(* IEC 61131-3 sources: 2026_Projet_YGO_ExcavatriceDragage/CODE/M_MAIN, 4 files *)

(* ---- GVL_Global.st ---- *)
(* ═══════════════════════════════════════════════════════════════
   🌐 GVL_Global — Variables globales d'utilité générale
   ───────────────────────────────────────────────────────────────
   🎯 Rôle : Horloges et signaux système partagés non persistants.
   📄 Docs : DOC/AF/AF_Partie-02_Architecture_Programme_v3.2.md
   ═══════════════════════════════════════════════════════════════ *)
{attribute 'qualified_only'}
VAR_GLOBAL
    BlinkClock                 : BOOL; // Horloge clignotement système (IHM/diag), rythme réglable GVL_PERSISTENT
END_VAR

(* ---- PRG_04_Treuils_Benne.st ---- *)
(* ═══════════════════════════════════════════════════════════════
   🪝 PRG_04_Treuils_Benne — Commande des Treuils M1 (moteur de retenue) / M2 (moteur Benne), Synchro et Benne
   ───────────────────────────────────────────────────────────────
   ⚙️ Exécuté par la tâche PLC en position 4 (après PRG_03_Modes_Cycle).
   ✅ Arbitre entre les commandes Manuelles (Joystick) et Automatiques (PRG_03_Modes_Cycle).
   📄 Docs : DOC/AF/AF_Partie-10_Fonction_Winch_v2.1.md ; DOC/AF/AF_Partie-10_Fonction_Winch/FB_Bucket_v1.0.md
   ═══════════════════════════════════════════════════════════════ *)

PROGRAM PRG_04_Treuils_Benne

VAR_INPUT
    // === 📥 ENTRÉES PROGRAMME (AUCUNE - PILOTÉ VIA PRG_02 & PRG_03) ===
END_VAR

VAR_OUTPUT
    // === 🚌 BUS INTER-PRG (producteur unique) ===
    Data : ST_WinchInterPrg; // <-- [BUS] Demandes finales, états, sécurités, synchro, benne
END_VAR

VAR
    instWinchSync : FB_WinchSync;
    instBucket   : FB_Bucket;
    // Seuil d'ouverture benne déclarant la fermeture atteinte (FB PUR). Instance PROPRE à
    // PRG_04 : l'arrivée de fermeture est évaluée DANS FB_Bucket, donc sur la mesure du
    // scan même, avant que PRG_04 ne puisse lire ses sorties. Les deux appels portent des
    // entrées identiques au même scan -> même décision, aucun critère dupliqué.
    instCloseThreshold : FB_BucketCloseThreshold;
    ThresholdMeasureValid : BOOL;  // Qualification de la mesure pour la branche seuil (références M1/M2 + défauts + référence benne)
    instSafetyWinchM1 : FB_Safety_Winch;   // Sécurité treuil M1 (SafeStop / permits / PowerCutOff)
    instSafetyWinchM2 : FB_Safety_Winch;
    instWinchM1   : FB_Winch;
    instWinchM2   : FB_Winch;
    // Projection lecture seule des états IHM treuils () : décharge la §8
    // (~250 lignes d'assignations pures) en un FB. Recopie bit-identique des
    // sources → WinchM1State/WinchM2State/WinchM1Safety/WinchM2Safety/CableLimitAscent.
    instWinchStateProjection : FB_WinchStateProjection;
    // Estimateurs bande vitesse réelle : alimentent le garde-fou palier FB_Winch
    // via MeasuredSpeedBand, 1 instance par treuil, mêmes sources que FB_Safety_Winch.
    instWinchLoadEstimatorM1 : FB_WinchLoadEstimator;
    instWinchLoadEstimatorM2 : FB_WinchLoadEstimator;

    // Collecteurs passifs d'apprentissage vitesse par palier : 1 par treuil,
    // écrivent la table RETAIN _WinchSpeedLearnTable {axe x sens x charge/vide x palier}.
    // STRICTEMENT PASSIFS : aucune commande moteur, aucune surveillance survitesse.
    instWinchSpeedLearningM1 : FB_WinchSpeedLearning;
    instWinchSpeedLearningM2 : FB_WinchSpeedLearning;
    // Dérivations des entrées de collecte (charge présente / conditions stables) — voir §6.
    LoadPresentM1 : BOOL;
    LoadPresentM2 : BOOL;
    StableForLearnM1 : BOOL;
    StableForLearnM2 : BOOL;

    // === FB D'ARBITRAGE DE COMMANDE (POO) ===
    instArbM1 : FB_WinchCmdArbitrationM1;  // * [INST] Arbitrage commande treuil M1
    instArbM2 : FB_WinchCmdArbitrationM2;  // * [INST] Arbitrage commande treuil M2
    instArbBucket : FB_BucketCmdArbitration;  // * [INST] Arbitrage commande benne (POO §5)

    // === REQUETES D'AXE ASSEMBLEES AVANT APPEL FB_WINCH ===
    // CODESYS n'accepte pas l'initialiseur de struct anonyme en parametre d'appel :
    // les structs WinchRequest / Sensors / Config sont remplies champ par champ ici.
    ReqM1Winch                   : ST_fbWinch_Req;             // . [LOC] Requête axe M1 (ordre, palier, bornes)
    ReqM2Winch                   : ST_fbWinch_Req;             // . [LOC] Requête axe M2 (ordre, palier, bornes)
    M1WinchSensors               : ST_fbWinch_Sensors;        // . [LOC] Mesures et feedbacks M1
    M2WinchSensors               : ST_fbWinch_Sensors;        // . [LOC] Mesures et feedbacks M2
    M1WinchCfg                   : ST_fbWinch_Cfg;            // . [LOC] Config statique M1 (table paliers, ralentissement)
    M2WinchCfg                   : ST_fbWinch_Cfg;            // . [LOC] Config statique M2 (table paliers, ralentissement)

    // === 📊 STRUCTS INTERNES (publiés via Data) ===
    WinchM1FinalInterlockRequest : ST_WinchFinalInterlockRequest; // . [LOC] Demande finale et interlocks treuil M1
    WinchM2FinalInterlockRequest : ST_WinchFinalInterlockRequest; // . [LOC] Demande finale et interlocks treuil M2
    KoboldContactorCmdArbitrated : BOOL;                         // . [LOC] Ordre contacteur capteur fond Kobold
    WinchM1State                 : ST_WinchState;                // . [LOC] Etat public treuil Retenue M1
    WinchM2State                 : ST_WinchState;                // . [LOC] Etat public treuil Benne M2
    WinchM1Safety                : ST_SafetyWinch;               // . [LOC] Diagnostic et securites treuil M1
    WinchM2Safety                : ST_SafetyWinch;               // . [LOC] Diagnostic et securites treuil M2
    SyncState                    : ST_SyncState;                 // . [LOC] Etat synchronisation treuils M1/M2
    BucketState                  : ST_BucketHMIState;            // . [LOC] Etat de fonctionnement benne
    Benne_IsRoughlyClosed        : BOOL;                         // . [LOC] Benne consideree fermee
    ArmingPermit                 : BOOL;                         // . [LOC] Permission d'armement homme-mort (combiné interlock benne, Option B)

    WinchBothMotionActive : BOOL;
    WinchBothMotionReady         : BOOL;                         // . [LOC] Verrou atomicite demarrage couple : les 2 treuils prets (hors dead-time D18, hors defaut latche)
    WinchBothFinalRequestsCoherent : BOOL;                       // . [LOC] Egalite effective des demandes physiques M1/M2 du scan
    WinchBothFinalStep45Coherent : BOOL;                         // . [LOC] Exception T291-A exacte : descente M1=P4 / M2=P5 en auto AX4..AX7
    WinchBothReqAscent           : BOOL;
    WinchBothReqDescend          : BOOL;
    ManualBottomPositionConfirmed  : BOOL;
    BottomPositionConfirmed        : BOOL;
    CmdBucketCloseArbitrated       : BOOL;

    // Séquencement automatique benne en pilotage both normal --
    // descente uniquement benne ouverte, montée uniquement benne
    // fermée. Distinct de DumpAtTremie/DiveSearch/ExtractionAssist (fonctionnement normal,
    // pas une assistance MAINT_N1/N2 dédiée). Réutilise WinchBothMotionActive/
    // WinchBothMotionDirection (§1 ci-dessus) : déjà exactement "mouvement both
    // demandé" dans les 2 modes (joystick Select=0, ou BtnWinchBothAscent/Descent) — mêmes variables
    // déjà utilisées par instBucket/instDiveSearch/instExtractionAssist.
    WinchBothDiveBucketOpenArmed     : BOOL;  // CmdOpen_IHM déclenché par ce mécanisme (diagnostic IHM)
    WinchBothMotionBlockedByBucket   : BOOL;  // Garde-fou direct -- voir §3
    WinchBothAscentBucketCloseArmed  : BOOL;  // CmdClose_IHM déclenché par ce mécanisme (diagnostic IHM)
    BucketBusyRiseEdge             : R_TRIG; // Détecte le début d'une action benne (Busy monté)
    BucketBusyFallEdge             : F_TRIG; // Détecte la fin d'une action benne (Busy retombé)
    ControlAscentArmedForThisClose : BOOL;   // Mémorise si LA fermeture en cours a été armée par ce mécanisme
    ExtractionControlActive        : BOOL;   // Phase vitesse contrôlée en cours (diagnostic IHM)
    ControlAscentStartM1PosM       : REAL;
    ControlAscentStartM2PosM       : REAL;

    // === ACTION BENNE M2 (bits directionnels, câblés au FB d'arbitrage) ===
    BucketM2ReqAscent  : BOOL;
    BucketM2ReqDescend : BOOL;
    M2AscentPermitApplied : BOOL;
    M2DescendPermitApplied : BOOL;

    // === STRUCTS D'ARBITRAGE (remplis champ par champ, CODESYS refuse l'init anonyme en appel) ===
    ArbIHM     : ST_fbWinchCmdArbitration_IHM;      // . [LOC] Entrées IHM FB d'arbitrage (partagé M1/M2)
    ArbContext : ST_fbWinchCmdArbitration_Context;  // . [LOC] Contexte gating FB d'arbitrage (partagé M1/M2)
    ArbM1Cfg   : ST_fbWinchCmdArbitration_Cfg;      // . [LOC] Config M1 (palier boutons/both)
    ArbM2Cfg   : ST_fbWinchCmdArbitration_Cfg;      // . [LOC] Config M2 (palier boutons/both + override benne)
    ArbBucketIHM     : ST_fbBucketCmdArbitration_IHM;      // . [LOC] Entrées IHM FB d'arbitrage benne
    ArbBucketContext : ST_fbBucketCmdArbitration_Context;  // . [LOC] Contexte gating FB d'arbitrage benne

    M1LogicRunRequest            : BOOL;
    M1LogicReqAscent             : BOOL;
    M1LogicReqDescend            : BOOL;
    M1LogicRequestStepTgt       : INT;   // Palier arbitré M1 (1..5, 0 = arrêt) — consommé par FB_Winch
    M1LogicRequestSpeedCmd_Pct  : REAL;  // Diagnostic % M1 (palier→%, IHM / simu)

    M2LogicRunRequest            : BOOL;
    M2LogicReqAscent             : BOOL;
    M2LogicReqDescend            : BOOL;
    M2LogicRequestStepTgt       : INT;   // Palier arbitré M2 (1..5, 0 = arrêt) — consommé par FB_Winch
    M2LogicRequestSpeedCmd_Pct  : REAL;  // Diagnostic % M2 (palier→%, IHM / simu)

    BottomLimitM1_Active    : REAL;
    BottomLimitM2_Active    : REAL;

    CableLimitAscentM1Reached : BOOL;
    CableLimitAscentM2Reached : BOOL;

    SafeStopM1_Raw          : BOOL;
    SafeStopM2_Raw          : BOOL;
    WinchContactorMismatchLvl1 : BOOL;   // . [LOC] niveau 1 : discordance contacteurs M1/M2 confirmee (amont OU vecteurs finaux) -> SafeStop
    SyncOperationPermit        : BOOL;   // . [LOC] Gate canonique : la surveillance d'ecart M1/M2 (synchro process + MecaE croise) est autorisee. FAUX pendant tout homing / toute manipulation benne.
    BucketActivityHold         : TOF;    // . [LOC] Maintien de la coupure surveillance synchro 4 s APRES la fin d'une action benne (transitoire d'arret treuils : coast + settle codeur -> faux ecart M1/M2)
    SafeStopM1_Active       : BOOL;
    SafeStopM2_Active       : BOOL;
    // Disponibilité de mouvement par axe/sens + conditions de base ArmingPermit
    ArmM1AscentAvail        : BOOL;
    ArmM1DescendAvail       : BOOL;
    ArmM2AscentAvail        : BOOL;
    ArmM2DescendAvail       : BOOL;
    ArmM3TremieAvail        : BOOL;
    ArmM3MaintenanceAvail   : BOOL;
    ArmAnyAxisAvail         : BOOL;
    ArmBucketBusy           : BOOL;
    ArmModeDisabled         : BOOL;
    ArmContactorOff         : BOOL;
    ArmPowerCutOff          : BOOL;
    // Taxonomie permit (D-P1 à D-P11) : SafetyPermit (safety pure), ProcessPermit (process pur),
    // ProcessAndSafetyPermit (= Safety AND Process), EffectivePermit (= couplage synchro).
    SafetyPermitM1_Descend   : BOOL;
    SafetyPermitM2_Descend   : BOOL;
    SafetyPermitM1_Ascent    : BOOL;
    SafetyPermitM2_Ascent    : BOOL;
    ProcessPermitM1_Descend  : BOOL;
    ProcessPermitM2_Descend  : BOOL;
    ProcessPermitM1_Ascent   : BOOL;
    ProcessPermitM2_Ascent   : BOOL;
    ProcessAndSafetyPermitM1_Descend : BOOL;
    ProcessAndSafetyPermitM2_Descend : BOOL;
    ProcessAndSafetyPermitM1_Ascent  : BOOL;
    ProcessAndSafetyPermitM2_Ascent  : BOOL;
    EffectivePermitM1_Descend : BOOL;
    EffectivePermitM2_Descend : BOOL;
    EffectivePermitM1_Ascent  : BOOL;
    EffectivePermitM2_Ascent  : BOOL;
    EffectivePermitBucket_Open  : BOOL;
    EffectivePermitBucket_Close : BOOL;

    // === 🔗 ATOMICITÉ BOTH — états agrégés explicites ===
    // CoupledBoth := couplage atomique M1/M2 indépendant de SyncEnable : actif en
    // synchro classique (anti-télescopage) OU dès qu'un mouvement both est demandé
    // (même si SyncEnable=FALSE en MAINT_N2). Une permission ou un SafeStop d'un
    // treuil bloque alors l'autre : départ jamais isolé.
    CoupledBoth             : BOOL;
    // Diagnostic IHM : Both bloqué + cause priorisée (voir §5).
    BothBlocked             : BOOL;
    BothBlockReason         : E_WinchTraceBlockReason;

    BenneBusyFallEdge     : F_TRIG;

    // Arrêt auto descente sur détection fond Kobold (pilotage normal)
    KoboldAutoStopRiseEdge  : R_TRIG;
    KoboldAutoStopFallEdge  : F_TRIG;
    KoboldImmersionConfirmed: BOOL;
    KoboldBottomTouchLatched: BOOL;
    DescendPermitDiveBucketOpen : BOOL; // mode Dive actif + benne ouverte = descente permise
    // pilotage unitaire M2 "sécurisé" -- bornes ouvert/fermé + palier 1
    ManualBucketLimitsActive : BOOL;
    ManualBucketJogActive    : BOOL; // WinchSel=2 + MAINT : jog benne unitaire M2 (ouv/ferm), indépendant du toggle bornes
    T248BucketJogActive : BOOL; // Phase JOG du séquencement benne-auto couplé (CoupledBucketPhaseLocked) : borne alignée sur l'état franc IsClosed/IsOpen, caduque dès Arbitrated=0
    M2JogApproachOpen        : BOOL; // M2 dans la zone de ralentissement avant l'arrêt ouverture (palier 1)
    M2JogApproachClose       : BOOL; // M2 dans la zone de ralentissement avant l'arrêt fermeture (palier 1)
    SlackCableAscentCapStep1    : BOOL; // mou de câble en récupération -- bride la montée au Palier 1
    BucketNotClosedAscentCapStep1 : BOOL; // benne non fermée à 100% à la montée -- bride la montée au Palier 1

    // Bypass simplifié séquence FB_DiveSearch -- front montant
    // Kobold pendant une descente couplée confirme directement le fond, sans passer par les
    // préconditions strictes de FB_DiveSearch (benne ouverte, DiveStartMin_M, fenêtre immersion).
    // FB_DiveSearch continue de tourner en parallèle (KoboldMeasureEnable toujours câblé
    // dessus) -- ce bypass est un chemin ADDITIONNEL, pas un remplacement.
    BypassKoboldFallEdge       : F_TRIG; // front descendant Kobold
    BypassKoboldBottomTouched  : BOOL;

    SyncMinorDeviation      : BOOL;
    SyncMinorDeviationBlocksUp   : BOOL;
    SyncMinorDeviationBlocksDown : BOOL;
    M2_LimitShift                : REAL;

    EffectiveMaxStepAscent    : INT;
    EffectiveMaxStepDescent  : INT;

    // Plafonds fixes de sécurité en position Maintenance (non réglables IHM).
    MaintenanceMaxStepAscent  : INT;
    MaintenanceMaxStepDescent : INT;

    // Agrégateur de clamp de palier — bornes communes M1=M2 puis M2-propre
    CommonMaxStepAscent   : INT;
    CommonMaxStepDescent : INT;
    CommonMinStepUp   : INT;
    CommonMinStepDown : INT;
    M2MaxStepUp       : INT;
    M2MaxStepDown     : INT;
    M2MinStepUp       : INT;
    M2MinStepDown     : INT;

    // Mémoire scan précédent pour SpeedDelta_Mps (IHM)
    M1_PrevSpeed_Mps : REAL;
    M2_PrevSpeed_Mps : REAL;

    // === MATRICE DE MAINTENANCE N1/N2 (AF-05 §4bis) ===
    // PRG_04 est le producteur unique du bypass EFFECTIF de son axe : FB_Safety_Winch / FB_Winch /
    // FB_Bucket ne connaissent que des booléens déjà gatés, jamais le mode (encapsulation AF03 §2).
    MaintN1 : BOOL;   // . [LOC] Mode MAINT_N1 arbitré (override FDC logiciel momentané)
    MaintN2 : BOOL;   // . [LOC] Mode MAINT_N2 arbitre (secours et pilotage direct contacteurs)
    ExtractionAssistActive : BOOL; // . [LOC] Séquence d'extraction active (mode MAINT + toggle) — gate permis de montée assistée

    // Override du FDC haut LOGICIEL — MAINT_N1, bouton IHM MAINTENU (jamais latché).
    // Le FDC haut CAPTEUR (TopPositionSensor ≈ 8,5 m) n'est JAMAIS ouvert par cet override.
    OverrideTopSoftwareN1M1 : BOOL;
    OverrideTopSoftwareN1M2 : BOOL;

    // Limite haute logicielle active (m) : 7,5 m nominal ➔ 8,5 m (capteur homing haut) sous override.
    TopLimitM1_M : REAL;
    TopLimitM2_M : REAL;

    // Bypass EFFECTIFS de la famille position (= bypass IHM armé, tous modes — dérogation MES 2026).
    // Servent au câblage ET à l'armement du re-homing obligatoire publié vers PRG_03 (PositionLimitOverriddenM1/M2).
    BypassM1TopLimitSwitchEff   : BOOL;
    BypassM1TopLimitSoftwareEff : BOOL;
    BypassM1CableLimitSwitchEff : BOOL;
    BypassM1LimitLegalEff       : BOOL;
    BypassM1MecaDEff            : BOOL;
    BypassM2TopLimitSwitchEff   : BOOL;
    BypassM2TopLimitSoftwareEff : BOOL;
    BypassM2CableLimitSwitchEff : BOOL;
    BypassM2LimitLegalEff       : BOOL;
    BypassM2MecaDEff            : BOOL;

    // Usage effectif d'un override/bypass de position -> arme le re-homing obligatoire (PRG_03).
    PositionLimitOverriddenM1 : BOOL;
    PositionLimitOverriddenM2 : BOOL;
    BrakeForceAllowedM1       : BOOL;
    BrakeForceAllowedM2       : BOOL;
    HomingFreeMoveBlockedN1   : BOOL;

    // 🕵️ Trace de blocage terrain (§8bis) — publiée via Data.TraceM1/M2, consommée FB_TroubleshootingView
    TraceM1               : ST_TraceWinch;        // . [LOC] Trace blocage treuil M1
    TraceM2               : ST_TraceWinch;        // . [LOC] Trace blocage treuil M2
    TraceM1_PrevReason    : E_WinchTraceBlockReason; // . [LOC] Cause précédente M1 (détection de changement)
    TraceM2_PrevReason    : E_WinchTraceBlockReason; // . [LOC] Cause précédente M2 (détection de changement)
END_VAR

{region "🎯 §1 Intention & assistants"}
// === 🪨 §1 INTENTION MAINTENANCE & ASSISTANTS ===

// Consommation de l'intention both continue opérateur (source unique PRG_03, tous modes)
WinchBothMotionActive    := PRG_03_Modes_Cycle.Data.WinchBothIntent.Active;
WinchBothReqAscent  := PRG_03_Modes_Cycle.Data.WinchBothIntent.ReqAscent;
WinchBothReqDescend := PRG_03_Modes_Cycle.Data.WinchBothIntent.ReqDescend;

// Récupération de l'état fond synthétisé par PRG_03
BottomPositionConfirmed := PRG_03_Modes_Cycle.Data.SequenceState.BottomTouchConfirmed;

// MODES DE MAINTENANCE (calculés en tête de scan : consommés dès §2 par instBucket)
// 🚨 DEROGATION MES septembre 2026 (AF-05 §4bis) : les bypass sécurité treuil M1/M2 + benne
// NE SONT PLUS conditionnés au mode. Un bypass IHM armé est effectif dans TOUS les modes
// (y compris SEMI_AUTO / AUTO). Choix opérateur assumé, tracé — voir AF-05 §4bis.
// MAINT_N1 reste utilisé pour l'override momentané du FDC haut logiciel (§5) et l'assistance extraction.
MaintN1 := (PRG_03_Modes_Cycle.Data.Auth.Mode = E_Mode.MAINT_N1);
MaintN2 := (PRG_03_Modes_Cycle.Data.Auth.Mode = E_Mode.MAINT_N2);
// Séquence d'extraction active (mode MAINT + toggle) : gate le permis de montée assistée (§5).
// Le permis lui-même (AscentPermit) est produit par FB_ExtractionAssist et consommé via le contrat benne.
// FB_ExtractionAssist retire (legacy, plus de toggle IHM) : gate desormais toujours ferme.
ExtractionAssistActive := FALSE;

// Jog benne unitaire M2 : joystick dédié M2 (WinchSel=2) en maintenance. Autorise
// l'ouverture (descente M2) hors mode Dive + active la détection passive d'état benne
// dans FB_Bucket. Indépendant du toggle bornes (TglManualBucketLimits).
ManualBucketJogActive := (PRG_03_Modes_Cycle.Data.Auth.JoystickWinchSelectArbitrated = 2)
    AND (PRG_03_Modes_Cycle.Data.Auth.Mode = E_Mode.MAINT_N1 OR PRG_03_Modes_Cycle.Data.Auth.Mode = E_Mode.MAINT_N2);

// Règle absolue en pilotage both normal --
// descente autorisée UNIQUEMENT benne ouverte, montée UNIQUEMENT benne fermée.
// Décision déléguée à FB_BucketCmdArbitration (POO §5) : flags armés + commandes
// arbitrées (ouverture, fermeture, contacteur Kobold). Bit-identique PRG_04 §1/§2.
ArbBucketIHM.BtnOpen  := GVL_IHM.M2TreuilBenne.Bucket.Cmd.BtnOpen;
ArbBucketIHM.BtnClose := GVL_IHM.M2TreuilBenne.Bucket.Cmd.BtnClose;

ArbBucketContext.TglEnableCoupledBucketSequencing := GVL_IHM.Commun.Cfg.TglEnableCoupledBucketSequencing
                                                    AND NOT PRG_02_Acquisition.Data.MachineHoming.Active;
ArbBucketContext.MotionActive   := WinchBothMotionActive;
ArbBucketContext.ReqAscent      := WinchBothReqAscent;
ArbBucketContext.ReqDescend     := WinchBothReqDescend;
ArbBucketContext.BucketIsOpen   := _BucketState.IsOpen;
ArbBucketContext.BucketIsClosed := _BucketState.IsClosed;
ArbBucketContext.CoupledPhaseLocked := PRG_03_Modes_Cycle.Data.Auth.CoupledBucketPhaseLocked;

instArbBucket(
    Enable    := NOT PRG_02_Acquisition.Data.MachineHoming.Active,
    Auth      := PRG_03_Modes_Cycle.Data.Auth,
    ReqBucket := PRG_03_Modes_Cycle.Data.ReqProgram.ReqBucket,
    IHM       := ArbBucketIHM,
    Context   := ArbBucketContext
);
WinchBothDiveBucketOpenArmed    := instArbBucket.WinchBothDiveBucketOpenArmed;
WinchBothAscentBucketCloseArmed := instArbBucket.WinchBothAscentBucketCloseArmed;
CmdBucketCloseArbitrated        := instArbBucket.CmdClose_IHM;
KoboldContactorCmdArbitrated    := instArbBucket.KoboldContactorCmdArbitrated;

{endregion}

{region "🪣 §2 Commande benne"}
// === 🏗️ §2 COMMANDE DU BENNE (FB_Bucket) ===

instBucket(
    Enable              := NOT PRG_03_Modes_Cycle.Data.Auth.InhibitM2,
    Reset               := PRG_07_Supervision.FaultMachineReset_IHM,
    PowerContactorEngaged     := PRG_02_Acquisition.HwIn.Machine.PowerContactorEngaged_DI,
    Mode                := PRG_03_Modes_Cycle.Data.Auth.Mode,
    CmdOpen_IHM         := instArbBucket.CmdOpen_IHM,
    CmdClose_IHM        := CmdBucketCloseArbitrated,
    // 🎛️ Seuil d'ouverture benne déclarant la fermeture atteinte. Réglage lu directement sur
    // GVL_IHM (patron déjà en place dans PRG_04 pour le plafond de montée contrôlée et la
    // distance de contrôle). Aucune copie locale : le FB clôt lui-même la plage, en défense
    // en profondeur.
    CloseReachedOpening_Pct := GVL_IHM.CycleSemiAuto.Cfg.ExtractionStartOpening_Pct,
    HoldAscentP1AfterClose := PRG_03_Modes_Cycle.Data.ReqProgram.ReqBucket.ReqHoldAscentP1AfterClose,
    ReqAscent           := WinchBothReqAscent OR (PRG_03_Modes_Cycle.Data.Auth.Mode = E_Mode.SEMI_AUTO AND PRG_02_Acquisition.Data.Joystick.AxisY.Direction > 0),
    ReqDescend          := WinchBothReqDescend OR (PRG_03_Modes_Cycle.Data.Auth.Mode = E_Mode.SEMI_AUTO AND PRG_02_Acquisition.Data.Joystick.AxisY.Direction < 0),
    EffectivePermitBucket_Open := EffectivePermitBucket_Open,
    EffectivePermitBucket_Close := EffectivePermitBucket_Close,
    CablePosM1          := PRG_02_Acquisition.Data.EncoderM1.Measurement.CablePosM,
    CablePosM2          := PRG_02_Acquisition.Data.EncoderM2.Measurement.CablePosM,
    HomedM1             := PRG_02_Acquisition.Data.EncoderM1.Homed,
    HomedM2             := PRG_02_Acquisition.Data.EncoderM2.Homed,
    HomedAndReliableM1  := PRG_02_Acquisition.Data.EncoderM1.HomedAndReliable,
    HomedAndReliableM2  := PRG_02_Acquisition.Data.EncoderM2.HomedAndReliable,
    HomingSuspectM1     := PRG_02_Acquisition.Data.EncoderM1.HomingSuspect,
    HomingSuspectM2     := PRG_02_Acquisition.Data.EncoderM2.HomingSuspect,
    WinchSelBucket      := (PRG_03_Modes_Cycle.Data.Auth.JoystickWinchSelectArbitrated = 2),
    BucketJogActive     := ManualBucketJogActive,
    ProgramBucketDriveActive := PRG_03_Modes_Cycle.Data.ReqProgram.ReqBucket.ReqOpen
                                OR PRG_03_Modes_Cycle.Data.ReqProgram.ReqBucket.ReqClose
                                OR PRG_03_Modes_Cycle.Data.ReqProgram.ReqBucket.ReqHoldAscentP1AfterClose,
    M1_Busy             := (instWinchM1.StepNumber > 0),
    M2_Busy             := (instWinchM2.StepNumber > 0),
    // Confirmations visuelles N2 : publication et offset benne. Le preset
    // materiel M2 associe est produit independamment dans PRG_02.
    ConfirmOpenPosition  := GVL_IHM.M2TreuilBenne.Bucket.Cmd.BtnConfirmOpenPos,
    ConfirmClosePosition := GVL_IHM.M2TreuilBenne.Bucket.Cmd.BtnConfirmClosePos,
    MachineHomingCommitOpen  := PRG_02_Acquisition.Data.MachineHoming.SetPosBucketOpen,
    MachineHomingCommitClose := PRG_02_Acquisition.Data.MachineHoming.SetPosBucketClose,
    InvalidateRef            := PRG_02_Acquisition.Data.MachineHoming.BucketRefInvalidate,
    MachineHomed := PRG_02_Acquisition.Data.MachineHoming.Homed,
    MachineHomingActive := PRG_02_Acquisition.Data.MachineHoming.Active,
    Config              := _BucketCfgPersist.Config,
    CfgTimeoutDuration     := GVL_IHM.M2TreuilBenne.Bucket.Cfg.CfgTimeoutDuration,
    BucketState        := _BucketState,
    InhibitM1           := PRG_03_Modes_Cycle.Data.Auth.InhibitM1,
    InhibitM2           := PRG_03_Modes_Cycle.Data.Auth.InhibitM2,
    // Bypass benne (n°25 de la matrice) — effectif tous modes si armé (dérogation MES 2026, AF-05 §4bis)
    BypassGlobal        := GVL_IHM.M2TreuilBenne.Bucket.Bypass.Global
);

// Auto-séquencement benne & Dégradation Palier 1
// Si la benne est en cours de fermeture/ouverture (instBucket.Busy), le mouvement couplé attend.
// Si la benne n'est pas fermée (NOT IsClosed) et que instBucket n'est plus occupé (Busy=FALSE),
// toute demande de montée est automatiquement dégradée au Palier 1 (Vitesse lente, voir instWinchM1/M2),
// protégeant ainsi la mécanique même en pilotage unitaire ou si l'auto-séquencement est désactivé.
// 📌 Note d'architecture (lag 1 scan) : M1/M2LogicRequestDirection est consommé ici avant son calcul arbitré
// en §3 (lag d'un cycle automate nominal, toléré et homogène avec les arbitrages Translation/Modes).
WinchBothMotionBlockedByBucket := WinchBothDiveBucketOpenArmed
                                 AND NOT instBucket.Lifecycle.Busy
                                 AND NOT PRG_02_Acquisition.Data.MachineHoming.Active;
BucketNotClosedAscentCapStep1 := NOT ManualBucketJogActive
    AND (M1LogicReqAscent OR M2LogicReqAscent)
    AND NOT instBucket.Lifecycle.Busy
    AND NOT _BucketState.IsClosed;

// === GATE CANONIQUE SURVEILLANCE ECART M1/M2 ===============================================
// REGLE MES : aucun defaut/alarme d'ecart M1/M2 (synchro process, MecaE croise, concordance
// contacteurs) ne doit apparaitre pendant un HOMING (machine ou codeur) ni pendant une
// MANIPULATION BENNE (auto Lifecycle.Busy OU jog unitaire) : dans ces phases M2-M1 varie
// volontairement jusqu'a ~15 m. Ce signal unique coupe la surveillance A LA SOURCE :
//   - instWinchSync.Enable
//   - instSafetyWinchM1/M2.CrossCheckEnable (latch MecaE)
//   - + FB_WinchSync purge ses latch a Enable=FALSE, + FB_Safety_Winch ouvre RefWindow sur
//     NOT CrossCheckEnable (RAZ continue MecaA/E).
// Tempo de RÉACTIVATION : 2 s après la fin d'une action benne (Lifecycle.Busy OU jog
// WinchSel=2), les treuils coastent encore et les codeurs se stabilisent -> l'écart
// serré 0,1 m de FB_WinchSync (SyncDeviationWarn, [SYNC] ErrorID:01) se déclenche à
// tort. Le TOF ne masque QUE FB_WinchSync (gate sur instWinchSync.Enable §4). MecaE
// croisé (tolérance ~2,5 m, absorbe le coast), MecaA et survitesse restent ACTIFS via
// CrossCheckEnable := SyncOperationPermit (inchangé) -> aucun trou de sécurité.
BucketActivityHold(IN := instBucket.Lifecycle.Busy
    OR ManualBucketJogActive
    OR GVL_IHM.M2TreuilBenne.Bucket.Cmd.BtnOpen
    OR GVL_IHM.M2TreuilBenne.Bucket.Cmd.BtnClose
    OR instArbBucket.CmdOpen_IHM
    OR instArbBucket.CmdClose_IHM
    OR PRG_03_Modes_Cycle.Data.ReqProgram.ReqBucket.ReqOpen
    OR PRG_03_Modes_Cycle.Data.ReqProgram.ReqBucket.ReqClose, PT := T#4s);

SyncOperationPermit := PRG_03_Modes_Cycle.Data.Auth.SyncEnable
    AND (PRG_03_Modes_Cycle.Data.Auth.JoystickWinchSelectArbitrated = 0)
    AND NOT PRG_02_Acquisition.Data.MachineHoming.Active
    AND NOT PRG_02_Acquisition.Data.EncoderM1.Measurement.HomingLifecycle.Busy
    AND NOT PRG_02_Acquisition.Data.EncoderM2.Measurement.HomingLifecycle.Busy
    AND NOT instBucket.Lifecycle.Busy
    AND NOT ManualBucketJogActive
    AND NOT GVL_IHM.M2TreuilBenne.Bucket.Cmd.BtnOpen
    AND NOT GVL_IHM.M2TreuilBenne.Bucket.Cmd.BtnClose
    AND NOT instArbBucket.CmdOpen_IHM
    AND NOT instArbBucket.CmdClose_IHM
    AND NOT PRG_03_Modes_Cycle.Data.ReqProgram.ReqBucket.ReqOpen
    AND NOT PRG_03_Modes_Cycle.Data.ReqProgram.ReqBucket.ReqClose
    // Pas de surveillance de synchronisme pendant les phases ou M1/M2 travaillent
    // volontairement de facon dissymetrique : contact fond, retente et fermeture/controle.
    // La surveillance est rearmee a partir de AX12 (montee en charge couplee).
    AND NOT (PRG_03_Modes_Cycle.Data.SequenceState.Step = E_AutoCycleStep.AX8_BOTTOM_CONFIRMED)
    AND NOT (PRG_03_Modes_Cycle.Data.SequenceState.Step = E_AutoCycleStep.AX9_RAISE_OFF_BOTTOM)
    AND NOT (PRG_03_Modes_Cycle.Data.SequenceState.Step = E_AutoCycleStep.AX10_CLOSE_BUCKET)
    AND NOT (PRG_03_Modes_Cycle.Data.SequenceState.Step = E_AutoCycleStep.AX11_CTRL_ASCENT)
    AND instBucket.ActiveOffsetValid;

// En mode récupération (SyncEnable=FALSE), si un mou de câble est détecté (bit3 ErrorId),
// la montée/enroulement est autorisée mais bridée au Palier 1 pour retendre le tambour en sécurité.
// 📌 Note d'architecture (lag 1 scan) : instSafetyWinchM1/M2.ErrorId est consommé ici avant l'exécution du FB
// au §5bis (lag d'un cycle automate nominal, sécurisé en amont par la lecture directe de M2_TensionedCable_DI).
SlackCableAscentCapStep1 := NOT GVL_IHM.Commun.Bypass.SlackCable
    AND NOT PRG_03_Modes_Cycle.Data.Auth.SyncEnable AND (
    ((instSafetyWinchM1.Fault.ErrorId AND 16#0008) <> 16#0000) OR
    ((instSafetyWinchM2.Fault.ErrorId AND 16#0008) <> 16#0000) OR
    (NOT PRG_02_Acquisition.HwIn.Winch.M2_TensionedCable_DI)
);

SyncMinorDeviation := (instWinchSync.Fault.ErrorId AND 16#0001) <> 16#0000;
// 🛡️ Soft-stop synchro : rattrapage directionnel volontaire UNIQUEMENT en
// commande unitaire. En commande BOTH (WinchBothMotionActive), l'écart mineur ne doit
// JAMAIS produire de rattrapage unilatéral d'un seul treuil — il est géré par le clamp
// palier §5ter (les 2 treuils sont bridés à 1) et le seuil critique (SafeStop des 2,
// §5). Donc les drapeaux sync sont coupés dès qu'un mouvement both est demandé.
SyncMinorDeviationBlocksUp   := _SyncSoftStopEnable AND SyncMinorDeviation AND (instWinchSync.SignedDeltaPosM > 0.0) AND NOT WinchBothMotionActive;
SyncMinorDeviationBlocksDown := _SyncSoftStopEnable AND SyncMinorDeviation AND (instWinchSync.SignedDeltaPosM < 0.0) AND NOT WinchBothMotionActive;

IF _CommunCfgPersist.WinchMaxStepAscent <= 0 THEN
    EffectiveMaxStepAscent := 5;
ELSE
    EffectiveMaxStepAscent := _CommunCfgPersist.WinchMaxStepAscent;
END_IF;

IF _CommunCfgPersist.WinchMaxStepDescent <= 0 THEN
    EffectiveMaxStepDescent := 5;
ELSE
    EffectiveMaxStepDescent := _CommunCfgPersist.WinchMaxStepDescent;
END_IF;

{endregion}

{region "🔀 §3 Arbitrage M1/M2"}
// === 🔀 §3 ARBITRAGE CONSIGNES M1 / M2 ===

// ── Arbitrage M1/M2 (FB_WinchCmdArbitrationM1/M2) ──
// Dérivation des bits d'action benne M2 (consommés par les 2 FB d'arbitrage)
BucketM2ReqAscent  := instBucket.M2_ReqAscent;
BucketM2ReqDescend := instBucket.M2_ReqDescend;

// Remplissage des structs d'arbitrage (champ par champ, CODESYS 3.5 refuse l'init anonyme en appel)
ArbIHM.BtnAscentM1           := GVL_IHM.M1TreuilRetenue.Cmd.BtnAscent;
ArbIHM.BtnDescentM1         := GVL_IHM.M1TreuilRetenue.Cmd.BtnDescent;
ArbIHM.BtnAscentM2           := GVL_IHM.M2TreuilBenne.Cmd.BtnAscent;
ArbIHM.BtnDescentM2         := GVL_IHM.M2TreuilBenne.Cmd.BtnDescent;
ArbIHM.BtnWinchBothAscent    := GVL_IHM.Commun.BtnWinchBothAscent;
ArbIHM.BtnWinchBothDescent  := GVL_IHM.Commun.BtnWinchBothDescent;

ArbContext.BucketBusy                     := instBucket.Lifecycle.Busy AND NOT MaintN2;
ArbContext.BucketM2RunRequest             := instBucket.M2_RunRequest AND NOT MaintN2;
ArbContext.BucketM2ReqAscent              := BucketM2ReqAscent;
ArbContext.BucketM2ReqDescend             := BucketM2ReqDescend;
ArbContext.BucketAutoCloseActive          := (PRG_03_Modes_Cycle.Data.Auth.Mode = E_Mode.SEMI_AUTO)
    AND (PRG_03_Modes_Cycle.Data.SequenceState.Step = E_AutoCycleStep.AX10_CLOSE_BUCKET)
    AND PRG_03_Modes_Cycle.Data.ReqProgram.ReqBucket.ReqClose;
ArbContext.BucketHandoffP1Active          := (PRG_03_Modes_Cycle.Data.Auth.Mode = E_Mode.SEMI_AUTO)
    AND (PRG_03_Modes_Cycle.Data.SequenceState.Step = E_AutoCycleStep.AX10B_RACCORDEMENT_P1)
    AND instBucket.CloseReached
    AND PRG_03_Modes_Cycle.Data.ReqProgram.ReqBucket.ReqHoldAscentP1AfterClose;
ArbContext.WinchBothMotionBlockedByBucket := WinchBothMotionBlockedByBucket AND NOT MaintN2;
ArbContext.SyncBlocksAscent                   := SyncMinorDeviationBlocksUp AND NOT MaintN2;
ArbContext.SyncBlocksDescent                 := SyncMinorDeviationBlocksDown AND NOT MaintN2;
// 🔗 Atomicité Both : agrégats consommés par la commande both (§5 calcule
// Both*Permit APRÈS §3 → lag 1 scan assumé au gate d'arbitre, documenté comme les
// autres gates lag-1 de PRG_04 ; l'enforcement même-scan est assuré par le routage
// §6 vers FB_Winch).
ArbContext.M1AscentAllowed  := EffectivePermitM1_Ascent;
ArbContext.M1DescendAllowed := EffectivePermitM1_Descend;
ArbContext.M2AscentAllowed  := EffectivePermitM2_Ascent;
ArbContext.M2DescendAllowed := EffectivePermitM2_Descend;
ArbContext.BothBlock         := BothBlocked;

ArbM1Cfg.BtnStepTgt := 5;
ArbM2Cfg.BtnStepTgt := 5;
ArbM2Cfg.BucketOverrideStepUpTgt   := LIMIT(1, _BucketCfgPersist.Config.MaxStepUp, 5);
ArbM2Cfg.BucketOverrideStepDownTgt := LIMIT(1, _BucketCfgPersist.Config.MaxStepDown, 5);
ArbM2Cfg.BucketAutoMaxStepUp       := LIMIT(1, GVL_IHM.CycleSemiAuto.Cfg.CtrlAscentMaxStep, 2);

// ── Arbitrage M1 (FB_WinchCmdArbitrationM1) ──
instArbM1(
    Enable     := TRUE,
    Joystick   := PRG_02_Acquisition.Data.Joystick,
    Auth       := PRG_03_Modes_Cycle.Data.Auth,
    ReqWinch   := PRG_03_Modes_Cycle.Data.ReqProgram.ReqWinchM1,
    BothIntent := PRG_03_Modes_Cycle.Data.WinchBothIntent,
    IHM        := ArbIHM,
    TglJoystickMaster := GVL_IHM.Modes.Cmd.TglJoystickMaster,
    Context    := ArbContext,
    Cfg        := ArbM1Cfg
);
M1LogicRunRequest := instArbM1.RunRequest;
M1LogicReqAscent  := instArbM1.ReqAscent;
M1LogicReqDescend := instArbM1.ReqDescend;
M1LogicRequestStepTgt := instArbM1.StepTgt;
// Diagnostic % (palier→%) pour IHM / simu — borne haute du palier arbitré.
IF (M1LogicRequestStepTgt >= 1) AND (M1LogicRequestStepTgt <= 5) THEN
    M1LogicRequestSpeedCmd_Pct := _WinchSpeedStepTable.StepThreshold_Pct[M1LogicRequestStepTgt];
ELSE
    M1LogicRequestSpeedCmd_Pct := 0.0;
END_IF;

// ── Arbitrage M2 (FB_WinchCmdArbitrationM2) ──
instArbM2(
    Enable     := TRUE,
    Joystick   := PRG_02_Acquisition.Data.Joystick,
    Auth       := PRG_03_Modes_Cycle.Data.Auth,
    ReqWinch   := PRG_03_Modes_Cycle.Data.ReqProgram.ReqWinchM2,
    BothIntent := PRG_03_Modes_Cycle.Data.WinchBothIntent,
    IHM        := ArbIHM,
    TglJoystickMaster := GVL_IHM.Modes.Cmd.TglJoystickMaster,
    Context    := ArbContext,
    Cfg        := ArbM2Cfg
);
M2LogicRunRequest := instArbM2.RunRequest;
M2LogicReqAscent  := instArbM2.ReqAscent;
M2LogicReqDescend := instArbM2.ReqDescend;
M2LogicRequestStepTgt := instArbM2.StepTgt;

// T248 — HOLD DE TRANSITION : changement de selecteur en cours -> requetes M1/M2 forcees
// a 0 (arret rampe normale) jusqu'a l'arret confirme des 2 treuils. Pas de hand-off en
// mouvement jog<->couple -> supprime l'a-coup. Le mouvement suivant redemarre de zero.
IF PRG_03_Modes_Cycle.Data.Auth.WinchSelTransitionHold THEN
    M1LogicRunRequest := FALSE; M1LogicReqAscent := FALSE; M1LogicReqDescend := FALSE; M1LogicRequestStepTgt := 0;
    M2LogicRunRequest := FALSE; M2LogicReqAscent := FALSE; M2LogicReqDescend := FALSE; M2LogicRequestStepTgt := 0;
END_IF;

// D1/D3/D4/D6 : blocage mouvements libres MAINT_N1 en Step 0 (tant que NOT Homed) + gating directionnel homing
HomingFreeMoveBlockedN1 := MaintN1
                           AND NOT PRG_02_Acquisition.Data.MachineHoming.Homed
                           AND NOT PRG_02_Acquisition.Data.MachineHoming.Active;
IF HomingFreeMoveBlockedN1 THEN
    M1LogicRunRequest := FALSE; M1LogicReqAscent := FALSE; M1LogicReqDescend := FALSE; M1LogicRequestStepTgt := 0;
    M2LogicRunRequest := FALSE; M2LogicReqAscent := FALSE; M2LogicReqDescend := FALSE; M2LogicRequestStepTgt := 0;
ELSIF PRG_02_Acquisition.Data.MachineHoming.Active THEN
    IF PRG_02_Acquisition.Data.MachineHoming.CmdWinchSelect = 2 THEN
        M1LogicRunRequest := FALSE; M1LogicReqAscent := FALSE; M1LogicReqDescend := FALSE; M1LogicRequestStepTgt := 0;
        M2LogicReqAscent  := M2LogicReqAscent  AND PRG_02_Acquisition.Data.MachineHoming.AllowAscent;
        M2LogicReqDescend := M2LogicReqDescend AND PRG_02_Acquisition.Data.MachineHoming.AllowDescend;
        M2LogicRunRequest := M2LogicRunRequest AND (M2LogicReqAscent OR M2LogicReqDescend);
    ELSIF PRG_02_Acquisition.Data.MachineHoming.CmdWinchSelect = 0 THEN
        M1LogicReqAscent  := M1LogicReqAscent  AND PRG_02_Acquisition.Data.MachineHoming.AllowAscent;
        M1LogicReqDescend := M1LogicReqDescend AND PRG_02_Acquisition.Data.MachineHoming.AllowDescend;
        M1LogicRunRequest := M1LogicRunRequest AND (M1LogicReqAscent OR M1LogicReqDescend);
        M2LogicReqAscent  := M2LogicReqAscent  AND PRG_02_Acquisition.Data.MachineHoming.AllowAscent;
        M2LogicReqDescend := M2LogicReqDescend AND PRG_02_Acquisition.Data.MachineHoming.AllowDescend;
        M2LogicRunRequest := M2LogicRunRequest AND (M2LogicReqAscent OR M2LogicReqDescend);
    ELSE
        M1LogicRunRequest := FALSE; M1LogicReqAscent := FALSE; M1LogicReqDescend := FALSE; M1LogicRequestStepTgt := 0;
        M2LogicRunRequest := FALSE; M2LogicReqAscent := FALSE; M2LogicReqDescend := FALSE; M2LogicRequestStepTgt := 0;
    END_IF;
END_IF;
// Diagnostic % (palier→%) pour IHM / simu — borne haute du palier arbitré.
IF (M2LogicRequestStepTgt >= 1) AND (M2LogicRequestStepTgt <= 5) THEN
    M2LogicRequestSpeedCmd_Pct := _WinchSpeedStepTable.StepThreshold_Pct[M2LogicRequestStepTgt];
ELSE
    M2LogicRequestSpeedCmd_Pct := 0.0;
END_IF;

// Front de fin d'action benne (F_TRIG conservé pour §3bis ArmingPermit et extraction control).
// L'arrêt forcé de fin d'action benne est désormais géré en interne par les FB d'arbitrage.
BenneBusyFallEdge(CLK := instBucket.Lifecycle.Busy);

// Après une fermeture benne armée PAR CE mécanisme
// (pas ExtractionAssist, qui a déjà sa propre phase CONTROL_ASCENT), la montée couplée qui
// enchaîne démarre en vitesse contrôlée (palier 1) sur ExtractionControlDistance_M avant de
// repasser en paliers normaux.
BucketBusyRiseEdge(CLK := instBucket.Lifecycle.Busy);
IF BucketBusyRiseEdge.Q THEN
    ControlAscentArmedForThisClose := WinchBothAscentBucketCloseArmed;
END_IF;
IF BucketBusyFallEdge.Q AND ControlAscentArmedForThisClose THEN
    ExtractionControlActive := TRUE;
    ControlAscentStartM1PosM := PRG_02_Acquisition.Data.EncoderM1.Measurement.CablePosM;
    ControlAscentStartM2PosM := PRG_02_Acquisition.Data.EncoderM2.Measurement.CablePosM;
END_IF;
IF ExtractionControlActive THEN
    IF (ABS(PRG_02_Acquisition.Data.EncoderM1.Measurement.CablePosM - ControlAscentStartM1PosM) >= GVL_IHM.CycleSemiAuto.Cfg.ExtractionControlDistance_M)
       AND (ABS(PRG_02_Acquisition.Data.EncoderM2.Measurement.CablePosM - ControlAscentStartM2PosM) >= GVL_IHM.CycleSemiAuto.Cfg.ExtractionControlDistance_M) THEN
        ExtractionControlActive := FALSE;         // Distance de contrôle parcourue : paliers normaux
    ELSIF NOT (WinchBothMotionActive AND WinchBothReqAscent) THEN
        ExtractionControlActive := FALSE;         // Ascending relâchée/interrompue : annule la phase
    END_IF;
END_IF;

{endregion}

{region "🛡️ §3bis ArmingPermit"}
// === 🛡️ §3bis ARMINGPERMIT (général — permis de mouvement) ===
// ArmingPermit = permission d'armement homme-mort (entrée FB_Joystick, consommée PRG_02).
// Règle générale : on ne peut armer QUE si au moins un axe (treuil M1/M2 ou translation M3)
// a un permis de mouvement effectif. Sinon, aucun mouvement n'est possible → armement inutile
// et trompeur (l'opérateur croit pouvoir bouger alors que tout est bloqué).
// Calcul déplacé après §5bis (où EffectivePermitM1/M2_Ascent/Descend sont disponibles).
// Combiné interlock benne conservé : interdit l'armement pendant une action benne
// (instBucket.Lifecycle.Busy) et 1 scan après (BenneBusyFallEdge.Q).
// Polarité positive (NC-100) : TRUE = armement autorisé.
{endregion}

{region "🔄 §4 Synchro M1/M2"}
// === 🔄 §4 SYNCHRONISATION M1 / M2 ===

instWinchSync(
    // Surveillance synchro (ecart position + concordance contacteurs) UNIQUEMENT en
    // pilotage couple. En unitaire M1 ou M2 (JoystickWinchSelectArbitrated <> 0) les
    // deux treuils sont volontairement independants : comparer M1/M2 declencherait un
    // faux ContactorMismatch (M2 commande seul, M1 non) -> SafeStop.
    // Gate canonique SyncOperationPermit (calcule §1) : homing OU benne -> surveillance
    // coupee A LA SOURCE. + ActiveOffsetSettled (transitoire de recalage offset) + inhibitions.
    Enable          := SyncOperationPermit
                        AND instBucket.ActiveOffsetSettled
                        AND NOT BucketActivityHold.Q
                        AND NOT PRG_03_Modes_Cycle.Data.Auth.InhibitM1 AND NOT PRG_03_Modes_Cycle.Data.Auth.InhibitM2,
    Reset           := PRG_07_Supervision.FaultMachineReset_IHM,
    Mode            := PRG_03_Modes_Cycle.Data.Auth.Mode,
    CablePosM1      := PRG_02_Acquisition.Data.EncoderM1.Measurement.CablePosM,
    CablePosM2      := PRG_02_Acquisition.Data.EncoderM2.Measurement.CablePosM,
    HomedAndReliableM1 := PRG_02_Acquisition.Data.EncoderM1.HomedAndReliable,
    HomedAndReliableM2 := PRG_02_Acquisition.Data.EncoderM2.HomedAndReliable,
    SyncEnable      := PRG_03_Modes_Cycle.Data.Auth.SyncEnable,
    CfgSyncToleranceM  := _SyncCfgPersist.CfgSyncTolerance_M,
    CfgSyncCriticalToleranceM := _SyncCfgPersist.CfgSyncCriticalTolerance_M,
    ActiveOffsetM   := instBucket.ActiveOffsetM,
    RelayFwdM1      := instWinchM1.RelayFwd,
    RelayFwdM2      := instWinchM2.RelayFwd,
    RelayRevM1      := instWinchM1.RelayRev,
    RelayRevM2      := instWinchM2.RelayRev,
    Contactor1_M1   := instWinchM1.Contactor1,
    Contactor1_M2   := instWinchM2.Contactor1,
    Contactor2_M1   := instWinchM1.Contactor2,
    Contactor2_M2   := instWinchM2.Contactor2,
    Contactor3_M1   := instWinchM1.Contactor3,
    Contactor3_M2   := instWinchM2.Contactor3,
    Contactor4_M1   := instWinchM1.Contactor4,
    Contactor4_M2   := instWinchM2.Contactor4,
    BypassGlobal    := GVL_IHM.M1M2Sync.Bypass.Global
                       OR GVL_IHM.M1TreuilRetenue.Bypass.Global
                       OR GVL_IHM.M2TreuilBenne.Bypass.Global
                       OR GVL_IHM.M1TreuilRetenue.Bypass.ContactorFeedback
                       OR GVL_IHM.M2TreuilBenne.Bypass.ContactorFeedback
                       OR GVL_IHM.M1TreuilRetenue.Bypass.Safety
                       OR GVL_IHM.M2TreuilBenne.Bypass.Safety
                       OR GVL_IHM.M1TreuilRetenue.Bypass.Process
                       OR GVL_IHM.M2TreuilBenne.Bypass.Process,
    DescentStep45Permit := PRG_03_Modes_Cycle.Data.AutoDiveM1Step4M2Step5Active,
    SpeedStepTable  := _WinchSpeedStepTable
);

// Pas de reconstruction de table M2 : le clamp §5ter (M2MaxStep* := 1) suffit
// — StepNumber ≤ 1 → seuls les états P1 sont commandés.
// M2 consomme directement _WinchSpeedStepTable (table normale).

{endregion}

{region "🔗 §5 Couplage & sécurités"}
// === 🛑 §5 COUPLAGE CROISÉ & SÉCURITÉS ===

// La limite légale (profondeur min. autorisée) doit elle aussi
// bénéficier du ralentissement progressif avant arrêt (comme la limite câble physique), pas juste
// un arrêt sec (DescendPermit). Comme les 2 limites bornent la même
// direction (descente), on alimente FB_Winch.BottomLimitM avec la PLUS RESTRICTIVE des deux
// (MAX de 2 valeurs négatives = celle la moins profonde = atteinte en premier) : le ralentissement
// (FB_Winch §"RALENTISSEMENT AUTOMATIQUE SUR BORDURES") s'enclenche alors sur la bonne limite,
// légale ou câble, sans dupliquer le mécanisme.
// M2 : la limite basse est comparee a CablePosM2 BRUTE cote FB_Winch -> on la decale de
// l'offset benne actif (idem M2_LimitShift cote haut). Benne fermee, M2 a deroule
// ~OffsetCloseM de plus que M1 : sans ce decalage la limite basse M2 se declenche
// ~15 m trop tot (REX MES 2026-09-04). ActiveOffsetM est continu (pente bornee).
IF _CommunCfgPersist.LimitLegalEnabled THEN
    BottomLimitM1_Active := MAX(_WinchM1CfgPersist.CfgCableLimitDescent_M, _CommunCfgPersist.LimitLegalDepthMinAllowed_M);
    BottomLimitM2_Active := MAX(_WinchM2CfgPersist.CfgCableLimitDescent_M, _CommunCfgPersist.LimitLegalDepthMinAllowed_M) + instBucket.ActiveOffsetM;
ELSE
    BottomLimitM1_Active := _WinchM1CfgPersist.CfgCableLimitDescent_M;
    BottomLimitM2_Active := _WinchM2CfgPersist.CfgCableLimitDescent_M + instBucket.ActiveOffsetM;
END_IF;

// 🩺 InputModuleFault (AF06 §3bis) : un module DI TOR hors service rend indisponibles
// les retours frein/thermique/contacteurs/fin de course des DEUX treuils (VH_0800END,
// Local_Digital_IO) — pas de granularité par treuil possible, donc SafeStop des DEUX.
// Perte d'une reference auparavant valide en mouvement : arret controle des
// deux treuils, sans PowerCutOff additionnel. Le cycle libere la demande
// seulement apres le composite d'arret mecanique confirme.
// Discordance contacteurs M1/M2 = niveau 1 (SafeStop) sans masque hexa.
//   - instWinchSync.ContactorMismatch : sur les requetes amont (FB_Winch).
//   - PRG_06_Outputs.Data.ContactorMismatch : sur les vecteurs PHYSIQUES finaux
//     (scan N-1, PRG_06 s'execute apres PRG_04). Escalade -> ExternalSyncEscalation ci-dessous.
WinchContactorMismatchLvl1 := instWinchSync.ContactorMismatch OR PRG_06_Outputs.Data.ContactorMismatch;
SafeStopM1_Raw      := WinchContactorMismatchLvl1 OR instBucket.M1SlipDetected OR PRG_02_Acquisition.Data.InputModules.Fault
                       OR PRG_02_Acquisition.Data.MachineHoming.HomingLoss;
SafeStopM2_Raw      := WinchContactorMismatchLvl1 OR PRG_02_Acquisition.Data.InputModules.Fault
                       OR PRG_02_Acquisition.Data.MachineHoming.HomingLoss;

// Surveillance Kobold descente normale (hors FB_DiveSearch)
// : signal HwIn.Machine.M1_M2_KoboldBottomTouch_DI (même que instDiveSearch §1).
KoboldAutoStopRiseEdge(CLK := PRG_02_Acquisition.HwIn.Machine.M1_M2_KoboldBottomTouch_DI);
KoboldAutoStopFallEdge(CLK := PRG_02_Acquisition.HwIn.Machine.M1_M2_KoboldBottomTouch_DI);

// Levée du verrou au neutre du joystick/boutons ou si toggle désactivé
IF PRG_02_Acquisition.Data.Joystick.AtNeutralXY OR NOT GVL_IHM.Commun.Cfg.TglEnableKoboldAutoStopDescent THEN
    KoboldImmersionConfirmed := FALSE;
    KoboldBottomTouchLatched := FALSE;
END_IF;

// WinchBothMotionActive requis : cette surveillance ne s'arme qu'en pilotage
// BOTH (Select=0), pas en pilotage unitaire M1 (où WinchBothMotionDirection reflète
// quand même l'axe joystick brut).
// Qualification immersion : front montant Kobold dans la fenêtre [ImmersionLower_M..ImmersionUpper_M]
IF GVL_IHM.Commun.Cfg.TglEnableKoboldAutoStopDescent
   AND WinchBothMotionActive
   AND WinchBothReqDescend
   AND _BucketState.IsOpen
   AND KoboldAutoStopRiseEdge.Q THEN
    IF (PRG_02_Acquisition.Data.EncoderM1.Measurement.CablePosM <= GVL_IHM.CycleSemiAuto.Cfg.ImmersionUpper_M)
       AND (PRG_02_Acquisition.Data.EncoderM1.Measurement.CablePosM >= GVL_IHM.CycleSemiAuto.Cfg.ImmersionLower_M)
       AND (PRG_02_Acquisition.Data.EncoderM2.Measurement.CablePosM <= GVL_IHM.CycleSemiAuto.Cfg.ImmersionUpper_M)
       AND (PRG_02_Acquisition.Data.EncoderM2.Measurement.CablePosM >= GVL_IHM.CycleSemiAuto.Cfg.ImmersionLower_M) THEN
        KoboldImmersionConfirmed := TRUE;
    END_IF;
END_IF;

// Détection fond : front descendant Kobold APRÈS immersion confirmée
IF KoboldAutoStopFallEdge.Q AND KoboldImmersionConfirmed THEN
    KoboldBottomTouchLatched := TRUE;
    KoboldImmersionConfirmed := FALSE;
END_IF;

// Autorisation directe et explicite issue de PRG_03 (DiveSearch / Cycle)
DescendPermitDiveBucketOpen := PRG_03_Modes_Cycle.Data.ReqProgram.ReqBucket.DescendPermitDiveBucketOpen;

// Le bypass arrête aussi la descente instantanément, même doctrine que le mécanisme
// KoboldBottomTouchLatched.
// Mode "pilotage unitaire M2 sécurisé" : bornes du JOG MANUEL, portée STRICTE = sélecteur
// arbitré sur M2 seul (Arbitrated=2) + toggle IHM, HORS phase JOG du séquencement benne-auto
// couplé (CoupledBucketPhaseLocked, qui passe aussi par Arbitrated=2 mais possède sa propre
// borne ci-dessous). Ne s'applique
// JAMAIS au pilotage couplé (Arbitrated=0, MAINT ou SEMI_AUTO) : ces mouvements ont leurs
// propres permis process (DescendPermitDiveBucketOpen, séquence auto) et le couplage atomique
// M1/M2 propagerait toute coupure M2 en blocage total des deux treuils. Ne passe PAS par
// instBucket (pas de CloseReq/OpenReq mémorisé, jogging libre) -- bornes directes ouvert/fermé
// (mêmes offsets que FB_Bucket, relatifs à la position réelle de M1) + palier 1 (voir
// instWinchM2 §6 plus bas).
ManualBucketLimitsActive := GVL_IHM.M2TreuilBenne.Bucket.Cmd.TglManualBucketLimits
    AND (PRG_03_Modes_Cycle.Data.Auth.JoystickWinchSelectArbitrated = 2)
    AND NOT PRG_03_Modes_Cycle.Data.Auth.CoupledBucketPhaseLocked
    AND PRG_02_Acquisition.Data.EncoderM1.HomedAndReliable
    AND PRG_02_Acquisition.Data.EncoderM2.HomedAndReliable
    AND NOT (PRG_02_Acquisition.Data.MachineHoming.SoftLimitsOff
             AND PRG_02_Acquisition.Data.MachineHoming.Active);

ProcessPermitM1_Descend := NOT (KoboldBottomTouchLatched OR BypassKoboldBottomTouched) AND DescendPermitDiveBucketOpen;
// Phase JOG du séquencement benne-auto couplé (CoupledBucketPhaseLocked ET Arbitrated=2) :
// borne alignée sur la frontière
// RÉELLE IsClosed/IsOpen (CoherenceLimitM, même seuil que FB_Bucket), jamais sur l'anticipation
// -- sans mouvement pour "coaster" le reste du trajet, une coupure à l'anticipation laisse un
// trou permanent avant l'état franc. Caduque automatiquement dès que Arbitrated repasse à 0
// (phase couplée) : ne bride jamais le mouvement couplé qui suit.
T248BucketJogActive := PRG_03_Modes_Cycle.Data.Auth.CoupledBucketPhaseLocked
    AND (PRG_03_Modes_Cycle.Data.Auth.JoystickWinchSelectArbitrated = 2);
// Ce chemin (pilotage unitaire M2, hors instBucket) applique l'anticipation d'inertie
// OpenAnticipationM/CloseAnticipationM (mêmes que FB_Bucket, réglables IHM) pour couvrir
// aussi le jog unitaire. L'ouverture benne (descente M2) est permise soit par le mode Dive
// (DescendPermitDiveBucketOpen), soit par le jog benne unitaire en maintenance
// (ManualBucketJogActive) — sinon la benne ne pourrait plus s'ouvrir en WinchSel=2.
ProcessPermitM2_Descend := NOT (KoboldBottomTouchLatched OR BypassKoboldBottomTouched)
    AND (DescendPermitDiveBucketOpen OR ManualBucketJogActive)
    AND NOT (ManualBucketLimitsActive AND (PRG_02_Acquisition.Data.EncoderM2.Measurement.CablePosM <= (PRG_02_Acquisition.Data.EncoderM1.Measurement.CablePosM + _BucketCfgPersist.Config.OffsetOpenM + _BucketCfgPersist.Config.OpenAnticipationM)))
    AND NOT (T248BucketJogActive AND (PRG_02_Acquisition.Data.EncoderM2.Measurement.CablePosM <= (PRG_02_Acquisition.Data.EncoderM1.Measurement.CablePosM + _BucketCfgPersist.Config.OffsetOpenM + _BucketCfgPersist.Config.CoherenceLimitM)));

// Permis process de montee : contrat extraction commun aux deux axes.
// M2 conserve l'anticipation de fermeture du pilotage benne unitaire, deja appliquee
// historiquement dans ProcessAndSafetyPermitM2_Ascent (refactor sans changement fonctionnel).
// Meme doctrine que la descente ci-dessus (T248BucketJogActive, CoherenceLimitM).
ProcessPermitM1_Ascent := NOT ExtractionAssistActive
    OR PRG_03_Modes_Cycle.Data.ReqProgram.ReqBucket.AscentPermit;
ProcessPermitM2_Ascent := (NOT ExtractionAssistActive
    OR PRG_03_Modes_Cycle.Data.ReqProgram.ReqBucket.AscentPermit)
    AND NOT (ManualBucketLimitsActive AND (PRG_02_Acquisition.Data.EncoderM2.Measurement.CablePosM >= (PRG_02_Acquisition.Data.EncoderM1.Measurement.CablePosM + _BucketCfgPersist.Config.OffsetCloseM - _BucketCfgPersist.Config.CloseAnticipationM)))
    AND NOT (T248BucketJogActive AND (PRG_02_Acquisition.Data.EncoderM2.Measurement.CablePosM >= (PRG_02_Acquisition.Data.EncoderM1.Measurement.CablePosM + _BucketCfgPersist.Config.OffsetCloseM - _BucketCfgPersist.Config.CoherenceLimitM)));

// Zone de ralentissement jog unitaire M2 : palier 1 forcé dans les JogSlowdownZoneM
// derniers mètres AVANT le point d'arrêt anticipé (Offset ± Anticipation). Le "1 m d'avant"
// est donc calculé sur la cible anticipée, pas sur l'offset brut, et suit tout réglage IHM.
M2JogApproachOpen := ManualBucketJogActive
    AND (PRG_02_Acquisition.Data.EncoderM2.Measurement.CablePosM
         <= (PRG_02_Acquisition.Data.EncoderM1.Measurement.CablePosM
             + _BucketCfgPersist.Config.OffsetOpenM
             + _BucketCfgPersist.Config.OpenAnticipationM
             + _BucketCfgPersist.Config.JogSlowdownZoneM));
M2JogApproachClose := ManualBucketJogActive
    AND (PRG_02_Acquisition.Data.EncoderM2.Measurement.CablePosM
         >= (PRG_02_Acquisition.Data.EncoderM1.Measurement.CablePosM
             + _BucketCfgPersist.Config.OffsetCloseM
             - _BucketCfgPersist.Config.CloseAnticipationM
             - _BucketCfgPersist.Config.JogSlowdownZoneM));

// Decalage de la limite haute logicielle M2 : la benne pend jusqu'a OffsetCloseM sous M1,
// donc en pilotage benne (WinchSel=2) OU si la benne est/va etre fermee, M2 doit avoir la
// marge de montee pour atteindre M1 + OffsetCloseM (pas seulement sa position courante).
// Le latch _BucketState.IsClosed n'est plus stale grace au fix A (§4a efface un latch
// contredit par la mesure). En etat indetermine (jamais latche), le terme WinchSel=2
// garantit quand meme la marge pendant l'operation benne.
// La marge (BIG) est donnee si la benne est/va etre fermee OU des que l'operateur
// SELECTIONNE le mode benne (select joystick BRUT = 2, avant meme l'arbitrage WinchSel) :
// M2 doit pouvoir monter jusqu'a M1 + OffsetCloseM pour fermer. Sinon (benne ouverte,
// M2 suit M1) la limite M2 = celle de M1. Le FDC haut PHYSIQUE reste la barriere dure
// (non bypassable, FB_Safety_Winch:528-531) independamment de cette limite soft.
// Le decalage de la limite M2 = l'offset benne ACTIF, point. Comparer CablePosM2 brute a
// (limite + M2_LimitShift) revient exactement a comparer la position M2 CORRIGEE
// (CablePosM2 - ActiveOffsetM) a la limite nominale - meme reference que M1. L'ancienne
// formule (M1 + OffsetCloseM + 1.5 - CfgCableLimitAscent) suivait M1 avec du retard et
// s'alignait mal selon l'etat benne -> faux declenchement "cable ascent limite" (REX MES
// 2026-09-04 : benne fermee, 15 m deroules, comparaison sur la brute). ActiveOffsetM est
// continu (pente bornee) et suit deja l'ouverture reelle.
M2_LimitShift := instBucket.ActiveOffsetM;

{endregion}

{region "🧮 §5-0 Matrice N1/N2"}
// === 🛡️ §5-0 MATRICE DE MAINTENANCE (AF-05 §4bis) ===
// 🚨 DEROGATION MES septembre 2026 : bypass_effectif := bypass_IHM (armé) — SANS conditionnement
// de mode. Un bypass IHM armé est effectif dans TOUS les modes, SEMI_AUTO et AUTO inclus.
// Écart assumé (Directive Machines / ISO 13849) : traçabilité IHM + doc AF-05 §4bis.
// L'override du FDC haut logiciel reste momentané et propre à MAINT_N1 (§ ci-dessous).

// --- Override FDC haut LOGICIEL (décision Q8) ---------------------------------------------
// MAINT_N1 + bouton IHM MAINTENU ➔ la limite logicielle passe de 7,5 m à la position du capteur
// de homing haut (8,5 m). Relâché ➔ retour à 7,5 m au cycle suivant (aucune mémorisation).
// ⛔ Cet override n'ouvre PAS BypassTopLimitSwitch : le capteur physique haut reste la butée
// dure — si TopPositionSensor retombe, AscentPermit tombe (FB_Safety_Winch §3) ➔ arrêt matériel.
// ⛔ Conditionné à Homed ET NON HomingSuspect : sans référence de position fiable, la butée
// logicielle de FB_Safety_Winch (§3) ET la zone de ralentissement de FB_Winch (§3) sont
// neutralisées — relever la limite dans ce cas ne laisserait QUE le capteur physique comme
// protection, approché à pleine vitesse. Sans référence, il n'y a pas de « dépassement
// contrôlé » : l'override est refusé, seul reste le bypass N2 (acte conscient, tracé).
OverrideTopSoftwareN1M1 := MaintN1
                           AND PRG_02_Acquisition.Data.EncoderM1.Homed
                           AND NOT PRG_02_Acquisition.Data.EncoderM1.HomingSuspect
                           AND GVL_IHM.M1TreuilRetenue.Cmd.BtnOverrideTopSoftware;
OverrideTopSoftwareN1M2 := MaintN1
                           AND PRG_02_Acquisition.Data.EncoderM2.Homed
                           AND NOT PRG_02_Acquisition.Data.EncoderM2.HomingSuspect
                           AND GVL_IHM.M2TreuilBenne.Cmd.BtnOverrideTopSoftware;

// --- Bypass EFFECTIFS de la famille position (individuel OR commun, SANS gate de mode — dérogation MES 2026) ---
BypassM1TopLimitSwitchEff   := (GVL_IHM.M1TreuilRetenue.Bypass.TopLimitSwitch   OR GVL_IHM.Commun.Bypass.TopLimitSwitch);
BypassM1TopLimitSoftwareEff := (GVL_IHM.M1TreuilRetenue.Bypass.TopLimitSoftware OR GVL_IHM.Commun.Bypass.TopLimitSoftware);
BypassM1CableLimitSwitchEff := (GVL_IHM.M1TreuilRetenue.Bypass.CableLimitSwitch OR GVL_IHM.Commun.Bypass.CableLimitSwitch);
BypassM1LimitLegalEff       := (GVL_IHM.M1TreuilRetenue.Bypass.LimitLegal       OR GVL_IHM.Commun.Bypass.LimitLegal);
BypassM1MecaDEff            := GVL_IHM.M1TreuilRetenue.Bypass.MecaD;
BypassM2TopLimitSwitchEff   := (GVL_IHM.M2TreuilBenne.Bypass.TopLimitSwitch      OR GVL_IHM.Commun.Bypass.TopLimitSwitch);
BypassM2TopLimitSoftwareEff := (GVL_IHM.M2TreuilBenne.Bypass.TopLimitSoftware    OR GVL_IHM.Commun.Bypass.TopLimitSoftware);
BypassM2CableLimitSwitchEff := (GVL_IHM.M2TreuilBenne.Bypass.CableLimitSwitch    OR GVL_IHM.Commun.Bypass.CableLimitSwitch);
BypassM2LimitLegalEff       := (GVL_IHM.M2TreuilBenne.Bypass.LimitLegal          OR GVL_IHM.Commun.Bypass.LimitLegal);
BypassM2MecaDEff            := GVL_IHM.M2TreuilBenne.Bypass.MecaD;

// --- Limite haute logicielle active -------------------------------------------------------
// Nominal 7,5 m (CfgCableLimitAscent_M) ; 8,5 m (CfgTopSensorPos_M) sous override N1 momentané
// ou bypass N2 latché du FDC logiciel. M2 conserve son décalage benne (M2_LimitShift) dans les
// deux cas : l'override ne modifie que l'assiette de référence, pas la géométrie M1/M2.
// Le seuil haut nominal est un arrêt immédiat (distance de ralentissement = 0 m).
// En override/bypass MAINT, seul le FDC haut matériel définit la borne : il reste non-bypassable.
TopLimitM1_M := SEL(OverrideTopSoftwareN1M1 OR BypassM1TopLimitSoftwareEff,
                    _CommunCfgPersist.CfgCableLimitAscent_M,
                    _WinchM1CfgPersist.CfgTopSensorPos_M);
TopLimitM2_M := SEL(OverrideTopSoftwareN1M2 OR BypassM2TopLimitSoftwareEff,
                    _CommunCfgPersist.CfgCableLimitAscent_M + M2_LimitShift,
                    _WinchM2CfgPersist.CfgTopSensorPos_M + M2_LimitShift);
// EXEMPTION jog benne seule (WinchSel=2) : la formule ci-dessus, une fois M2_LimitShift
// applique, revient exactement a tester la position REELLE de M1 (M2_raw - ActiveOffsetM
// = M1). Resultat : quand M1 est deja au-dessus de CfgCableLimitAscent_M, fermer/ouvrir
// la benne (M2 seul, M1 IMMOBILE) est bloque par la meme limite que la montee de M1,
// alors que manipuler la benne ne fait jamais monter l'ensemble plus haut que M1 courant
// (REX MES 2026-09-04 : "le treuil ne change pas d'altimetrie en mvt benne"). En jog
// benne pur, on remplace donc la butee ALTITUDE ABSOLUE par une butee GEOMETRIQUE relative
// a M1 courant (OffsetCloseM + marge) : c'est deja le vrai limiteur mecanique de la benne
// (ManualBucketLimitsActive/anticipation, PRG_04 ~710-735). Le FdC haut MATERIEL
// (TopPositionSensor, FB_Safety_Winch) reste une barriere INDEPENDANTE et non affectee.
IF ManualBucketJogActive
   AND PRG_02_Acquisition.Data.EncoderM1.HomedAndReliable
   AND PRG_02_Acquisition.Data.EncoderM2.HomedAndReliable THEN
    TopLimitM2_M := PRG_02_Acquisition.Data.EncoderM1.Measurement.CablePosM
                     + _BucketCfgPersist.Config.OffsetCloseM + 2.0;
ELSIF WinchBothMotionActive AND NOT (OverrideTopSoftwareN1M2 OR BypassM2TopLimitSoftwareEff) THEN
    // En Both (WinchBothMotionActive), M1 est l'autorité nominale de montée et
    // d'arrêt haut. M2 devient un garde-fou dérivé avec marge de tolérance +0.50 m sur le FDC
    // logiciel haut pour éliminer les arrêts prématurés sur benne intermédiaire (réserve TOP >= 1.00 m respectée).
    TopLimitM2_M := _CommunCfgPersist.CfgCableLimitAscent_M + M2_LimitShift + 0.50;
END_IF;

// --- Usage effectif d'un override/bypass de position → re-homing obligatoire ---------------
// Publié vers PRG_03 (rang 03) ➔ FB_Modes arme HomingRequiredMx à la sortie du mode maintenance.
// Famille position : TopLimitSwitch, TopLimitSoftware, CableLimitSwitch, LimitLegal, MecaD
// (+ l'override N1 momentané).
PositionLimitOverriddenM1 := OverrideTopSoftwareN1M1 OR BypassM1TopLimitSwitchEff
                             OR BypassM1TopLimitSoftwareEff OR BypassM1CableLimitSwitchEff
                             OR BypassM1LimitLegalEff OR BypassM1MecaDEff;
PositionLimitOverriddenM2 := OverrideTopSoftwareN1M2 OR BypassM2TopLimitSwitchEff
                             OR BypassM2TopLimitSoftwareEff OR BypassM2CableLimitSwitchEff
                             OR BypassM2LimitLegalEff OR BypassM2MecaDEff;
{endregion}

{region "🛡️ §5bis Sécurité M1/M2"}

// FB_Safety_Winch M1/M2.
// Instancié avant instWinchM1/M2 : MovementCommanded lit RelayFwd/RelayRev du scan précédent
// (même lag 1 scan accepté que M4/Translation, jamais sur Reset/SafeStop/PowerCutOff/sortie finale).
BrakeForceAllowedM1 := MaintN2
    AND PRG_02_Acquisition.HwIn.Machine.EmergencyChainClosed_DI
    AND PRG_02_Acquisition.HwIn.Machine.PowerContactorEngaged_DI
    AND (GVL_IHM.MaintenanceN2.Cmd.BtnBothBrakeRelease OR GVL_IHM.MaintenanceN2.Cmd.BtnM1BrakeRelease);
BrakeForceAllowedM2 := MaintN2
    AND PRG_02_Acquisition.HwIn.Machine.EmergencyChainClosed_DI
    AND PRG_02_Acquisition.HwIn.Machine.PowerContactorEngaged_DI
    AND (GVL_IHM.MaintenanceN2.Cmd.BtnBothBrakeRelease OR GVL_IHM.MaintenanceN2.Cmd.BtnM2BrakeRelease);

instSafetyWinchM1(
    Enable                 := (PRG_03_Modes_Cycle.Data.Auth.Mode <> E_Mode.DISABLE) AND NOT PRG_03_Modes_Cycle.Data.Auth.InhibitM1,
    Reset                  := PRG_07_Supervision.FaultMachineReset_IHM,
    PowerContactorEngaged  := PRG_02_Acquisition.HwIn.Machine.PowerContactorEngaged_DI,
    Mode                   := PRG_03_Modes_Cycle.Data.Auth.Mode,
    SyncEnable             := PRG_03_Modes_Cycle.Data.Auth.SyncEnable,
    CrossCheckEnable       := SyncOperationPermit,
    JoystickOnline         := PRG_02_Acquisition.Data.Network.Joystick.Online,
    JoystickOperational    := PRG_02_Acquisition.Data.Network.Joystick.Operational,
    HeartbeatIhmOk         := GVL_IHM.Commun.HeartbeatIhmOk,
    EncoderAvailable       := PRG_02_Acquisition.Data.EncoderM1.Measurement.EncoderAvailable,
    EncoderFaultBypass     := GVL_IHM.M1TreuilRetenue.Bypass.EncoderFault,
    ThermalFeedback        := NOT PRG_02_Acquisition.HwIn.Winch.M1_ThermalOk_DI,
    BrakeThermalFeedback   := NOT PRG_02_Acquisition.HwIn.Machine.M1_M2_M3_BrakeThermalOk_DI,
    SlackCableDetected     := NOT PRG_02_Acquisition.HwIn.Winch.M2_TensionedCable_DI,
    PhaseRotationOk        := PRG_02_Acquisition.HwIn.Machine.PhaseRotationOk_DI,
    // FB_Safety_Winch attend le contact NC : TRUE = circuit sain / FdC haut libre.
    // FALSE = FdC haut atteint ou rupture de chaîne ; le FB bloque alors la montée.
    TopPositionSensor      := PRG_02_Acquisition.HwIn.Winch.M1M2_TopPositionFree_DI,
    InReferencingMode      := PRG_02_Acquisition.Data.EncoderM1.Measurement.HomingLifecycle.Busy,
    SoftLimitsBypassed     := PRG_02_Acquisition.Data.MachineHoming.SoftLimitsOff
                              AND PRG_02_Acquisition.Data.MachineHoming.Active,
    BrakeForceAllowed      := BrakeForceAllowedM1,
    CablePosM              := PRG_02_Acquisition.Data.EncoderM1.Measurement.CablePosM,
    CfgCableLimitDescentM  := _WinchM1CfgPersist.CfgCableLimitDescent_M,
    LimitLegalReached      := GVL_IHM.Commun.LimitLegalReached,
    ReqAscent              := M1LogicReqAscent,
    ReqDescend             := M1LogicReqDescend,
    MovementCommanded      := instWinchM1.RelayFwd OR instWinchM1.RelayRev,
    Homed                  := PRG_02_Acquisition.Data.EncoderM1.Homed,
    HomingSuspect          := PRG_02_Acquisition.Data.EncoderM1.HomingSuspect,
    TopLimitM              := TopLimitM1_M,
    FwdRevSpeedFeedbackOff := PRG_02_Acquisition.HwIn.Winch.M1_ContactorsReleased_DI,
    BrakeFeedback          := PRG_02_Acquisition.HwIn.Winch.M1_BrakeIsOpen_DI,
    JoystickYNeutral       := (PRG_02_Acquisition.Data.Joystick.AxisY.Direction = 0),
    BenneHoldStillActive   := instBucket.Lifecycle.Busy,
    ExpectedOtherWinchPosM := PRG_02_Acquisition.Data.EncoderM2.Measurement.CablePosM - instBucket.ActiveOffsetM,
    BenneBusy              := instBucket.Lifecycle.Busy,
    OtherWinchInhibited    := PRG_03_Modes_Cycle.Data.Auth.InhibitM2,
    MeasuredSpeedMps       := PRG_02_Acquisition.Data.EncoderM1.Measurement.Speed_Mps,
    MeasuredSpeedSignedMps := PRG_02_Acquisition.Data.EncoderM1.Measurement.SignedSpeed_Mps,
    MeasuredSpeedValid     := PRG_02_Acquisition.Data.EncoderM1.Measurement.SpeedValid,
    SpeedBandMaxMps        := _WinchSpeedConfig.SpeedBandMaxMps[5],
    // Matrice AF-05 §4bis : bypass transmis SANS gate de mode (dérogation MES 2026, tous modes).
    // Le bypass commun reste en OR avec l'individuel (pilotage "both") — câblage d'origine inchangé.
    BypassGlobal           := GVL_IHM.M1TreuilRetenue.Bypass.Global,
    BypassSafety           := GVL_IHM.M1TreuilRetenue.Bypass.Safety,
    BypassProcess          := (GVL_IHM.M1TreuilRetenue.Bypass.Process
                              OR GVL_IHM.Commun.Bypass.SlackCable),
    // OR avec le bypass commun (Commun.Bypass) -- leve la
    // protection sur les 2 treuils simultanement pour le pilotage "both", sans retirer le
    // bypass individuel pour le pilotage a l'unite.
    BypassTopLimitSwitch   := BypassM1TopLimitSwitchEff,
    BypassTopLimitSoftware := BypassM1TopLimitSoftwareEff,
    BypassCableLimitSwitch := BypassM1CableLimitSwitchEff,
    BypassLimitLegal       := BypassM1LimitLegalEff,
    BypassOperatorComm     := GVL_IHM.M1TreuilRetenue.Bypass.OperatorComm,
    BypassPhaseRotation    := GVL_IHM.M1TreuilRetenue.Bypass.PhaseRotation,
    BypassBrakeThermal     := GVL_IHM.M1TreuilRetenue.Bypass.BrakeThermal,
    BypassMotorThermal     := GVL_IHM.M1TreuilRetenue.Bypass.MotorThermal,
    BypassMecaA            := GVL_IHM.M1TreuilRetenue.Bypass.MecaA,
    BypassMecaB            := GVL_IHM.M1TreuilRetenue.Bypass.MecaB,
    BypassMecaC            := GVL_IHM.M1TreuilRetenue.Bypass.MecaC,
    BypassMecaD            := BypassM1MecaDEff,
    BypassMecaE            := GVL_IHM.M1TreuilRetenue.Bypass.MecaE,
    CriticalSyncToleranceM := _WinchCriticalSyncTolerance_M,
    ExternalSyncEscalation := PRG_06_Outputs.Data.ContactorMismatchEscalated,
    TopHardStopLatched     := PRG_06_Outputs.Data.TopHardStopLatched
);

instSafetyWinchM2(
    Enable                 := (PRG_03_Modes_Cycle.Data.Auth.Mode <> E_Mode.DISABLE) AND NOT PRG_03_Modes_Cycle.Data.Auth.InhibitM2,
    Reset                  := PRG_07_Supervision.FaultMachineReset_IHM,
    PowerContactorEngaged  := PRG_02_Acquisition.HwIn.Machine.PowerContactorEngaged_DI,
    Mode                   := PRG_03_Modes_Cycle.Data.Auth.Mode,
    SyncEnable             := PRG_03_Modes_Cycle.Data.Auth.SyncEnable,
    // Ecart critique croise M1/M2 (Meca E, FB_Safety_Winch:354) : gate canonique
    // SyncOperationPermit (homing/benne -> OFF). N'affecte PAS le routage mou-de-cable
    // (:508/:520) qui reste sur SyncEnable brut. Le mouvement couple par boutons-both
    // (WinchBothMotionActive sans WinchSel=0) est un cas residuel -> voir T-tache.
    CrossCheckEnable       := SyncOperationPermit,
    JoystickOnline         := PRG_02_Acquisition.Data.Network.Joystick.Online,
    JoystickOperational    := PRG_02_Acquisition.Data.Network.Joystick.Operational,
    HeartbeatIhmOk         := GVL_IHM.Commun.HeartbeatIhmOk,
    EncoderAvailable       := PRG_02_Acquisition.Data.EncoderM2.Measurement.EncoderAvailable,
    EncoderFaultBypass     := GVL_IHM.M2TreuilBenne.Bypass.EncoderFault,
    ThermalFeedback        := NOT PRG_02_Acquisition.HwIn.Winch.M2_ThermalOk_DI,
    BrakeThermalFeedback   := NOT PRG_02_Acquisition.HwIn.Machine.M1_M2_M3_BrakeThermalOk_DI,
    SlackCableDetected     := NOT PRG_02_Acquisition.HwIn.Winch.M2_TensionedCable_DI,
    PhaseRotationOk        := PRG_02_Acquisition.HwIn.Machine.PhaseRotationOk_DI,
    // Même contact NC que M1 : TRUE = FdC haut libre, FALSE = FdC atteint/chaîne ouverte.
    TopPositionSensor      := PRG_02_Acquisition.HwIn.Winch.M1M2_TopPositionFree_DI,
    InReferencingMode      := PRG_02_Acquisition.Data.EncoderM2.Measurement.HomingLifecycle.Busy,
    SoftLimitsBypassed     := PRG_02_Acquisition.Data.MachineHoming.SoftLimitsOff
                              AND PRG_02_Acquisition.Data.MachineHoming.Active,
    BrakeForceAllowed      := BrakeForceAllowedM2,
    CablePosM              := PRG_02_Acquisition.Data.EncoderM2.Measurement.CablePosM,
    CfgCableLimitDescentM  := _WinchM2CfgPersist.CfgCableLimitDescent_M,
    LimitLegalReached      := GVL_IHM.Commun.LimitLegalReached,
    ReqAscent              := M2LogicReqAscent,
    ReqDescend             := M2LogicReqDescend,
    MovementCommanded      := instWinchM2.RelayFwd OR instWinchM2.RelayRev,
    Homed                  := PRG_02_Acquisition.Data.EncoderM2.Homed,
    HomingSuspect          := PRG_02_Acquisition.Data.EncoderM2.HomingSuspect,
    TopLimitM              := TopLimitM2_M,
    FwdRevSpeedFeedbackOff := PRG_02_Acquisition.HwIn.Winch.M2_ContactorsReleased_DI,
    BrakeFeedback          := PRG_02_Acquisition.HwIn.Winch.M2_BrakeIsOpen_DI,
    JoystickYNeutral       := (PRG_02_Acquisition.Data.Joystick.AxisY.Direction = 0),
    BenneHoldStillActive   := FALSE,
    ExpectedOtherWinchPosM := PRG_02_Acquisition.Data.EncoderM1.Measurement.CablePosM + instBucket.ActiveOffsetM,
    BenneBusy              := instBucket.Lifecycle.Busy,
    OtherWinchInhibited    := PRG_03_Modes_Cycle.Data.Auth.InhibitM1,
    MeasuredSpeedMps       := PRG_02_Acquisition.Data.EncoderM2.Measurement.Speed_Mps,
    MeasuredSpeedSignedMps := PRG_02_Acquisition.Data.EncoderM2.Measurement.SignedSpeed_Mps,
    MeasuredSpeedValid     := PRG_02_Acquisition.Data.EncoderM2.Measurement.SpeedValid,
    SpeedBandMaxMps        := _WinchSpeedConfig.SpeedBandMaxMps[5],
    // Matrice AF-05 §4bis (identique à M1 ci-dessus)
    BypassGlobal           := GVL_IHM.M2TreuilBenne.Bypass.Global,
    BypassSafety           := GVL_IHM.M2TreuilBenne.Bypass.Safety,
    BypassProcess          := (GVL_IHM.M2TreuilBenne.Bypass.Process
                              OR GVL_IHM.Commun.Bypass.SlackCable),
    // OR avec le bypass commun (Commun.Bypass) -- voir M1 ci-dessus
    BypassTopLimitSwitch   := BypassM2TopLimitSwitchEff,
    BypassTopLimitSoftware := BypassM2TopLimitSoftwareEff,
    BypassCableLimitSwitch := BypassM2CableLimitSwitchEff,
    BypassLimitLegal       := BypassM2LimitLegalEff,
    BypassOperatorComm     := GVL_IHM.M2TreuilBenne.Bypass.OperatorComm,
    BypassPhaseRotation    := GVL_IHM.M2TreuilBenne.Bypass.PhaseRotation,
    BypassBrakeThermal     := GVL_IHM.M2TreuilBenne.Bypass.BrakeThermal,
    BypassMotorThermal     := GVL_IHM.M2TreuilBenne.Bypass.MotorThermal,
    BypassMecaA            := GVL_IHM.M2TreuilBenne.Bypass.MecaA,
    BypassMecaB            := GVL_IHM.M2TreuilBenne.Bypass.MecaB,
    BypassMecaC            := GVL_IHM.M2TreuilBenne.Bypass.MecaC,
    BypassMecaD            := BypassM2MecaDEff,
    BypassMecaE            := GVL_IHM.M2TreuilBenne.Bypass.MecaE,
    CriticalSyncToleranceM := _WinchCriticalSyncTolerance_M,
    ExternalSyncEscalation := PRG_06_Outputs.Data.ContactorMismatchEscalated,
    TopHardStopLatched     := PRG_06_Outputs.Data.TopHardStopLatched
);

SafeStopM1_Raw := SafeStopM1_Raw OR instSafetyWinchM1.SafeStop;
SafeStopM2_Raw := SafeStopM2_Raw OR instSafetyWinchM2.SafeStop;
// SafetyPermit = sorties FB_Safety_Winch (safety pure)
SafetyPermitM1_Descend := instSafetyWinchM1.DescendPermit;
SafetyPermitM2_Descend := instSafetyWinchM2.DescendPermit;
SafetyPermitM1_Ascent  := instSafetyWinchM1.AscentPermit;
SafetyPermitM2_Ascent  := instSafetyWinchM2.AscentPermit;
// ProcessAndSafetyPermit = Safety AND Process (ex _Raw)
ProcessAndSafetyPermitM1_Descend := ProcessPermitM1_Descend AND SafetyPermitM1_Descend;
ProcessAndSafetyPermitM2_Descend := ProcessPermitM2_Descend AND SafetyPermitM2_Descend;

// Mode "vidage à la trémie" : descente M1 interdite tant que M3 n'est pas à P1 (travail)
// ou en position Maintenance -- verrouille la descente-treuil (payout cable reel) / la
// translation, pour se rapprocher d'un enchaînement automatique sûr.
// M2 EXEMPTE quand seule la benne bouge (jog unitaire WinchSel=2 ou programme benne) :
// ouvrir/fermer la benne (M2 seul, M1 immobile) N'EST PAS une descente treuil verticale
// -> ça doit rester possible a la Tremie (design d'origine : "a la Tremie, seul open/close
// benne permis"). Sans cette exemption, EffectivePermitBucket_Open/Close (cable sur
// EffectivePermitM2_Descend/Ascent, ligne ~1004) heritait du meme verrou par accident de
// cablage -> ouverture benne bloquee a la Tremie (REX MES 2026-09-04).
// Décision et calcul centralisés dans PRG_03_Modes_Cycle.Data.SequenceState.WinchDescentAuth_M3
IF NOT PRG_03_Modes_Cycle.Data.SequenceState.WinchDescentAuth_M3 THEN
    ProcessAndSafetyPermitM1_Descend := FALSE;
    IF NOT (ManualBucketJogActive
            OR PRG_03_Modes_Cycle.Data.ReqProgram.ReqBucket.ReqOpen
            OR PRG_03_Modes_Cycle.Data.ReqProgram.ReqBucket.ReqClose) THEN
        ProcessAndSafetyPermitM2_Descend := FALSE;
    END_IF;
END_IF;
// Permis de montée assistée : consommé depuis FB_ExtractionAssist (via le contrat benne).
// Hors extraction (NOT ExtractionAssistActive), la montée reste libre ; pendant l'extraction,
// la montée n'est autorisée que si l'assistant la délivre (AscentPermit, qui intègre les
// conditions process AscentControlSafe/AscentNominalSafe). Polarité fail-safe (TRUE = autorisé).
ProcessAndSafetyPermitM1_Ascent := ProcessPermitM1_Ascent AND SafetyPermitM1_Ascent;
ProcessAndSafetyPermitM2_Ascent := ProcessPermitM2_Ascent AND SafetyPermitM2_Ascent;

// 🔗 Couplage atomique M1/M2 : indépendant de SyncEnable. Actif en synchro
// classique (anti-télescopage) OU dès qu'un mouvement both est demandé — même si
// SyncEnable=FALSE (ex. MAINT_N2). Permet qu'une permission ou un SafeStop d'un
// treuil bloque l'autre : départ jamais isolé. WinchBothMotionActive est défini en
// §1 (disponible avant §5).
CoupledBoth := instWinchSync.SyncActive OR WinchBothMotionActive;

SafeStopM1_Active := SafeStopM1_Raw OR (CoupledBoth AND SafeStopM2_Raw);
SafeStopM2_Active := SafeStopM2_Raw OR (CoupledBoth AND SafeStopM1_Raw);
// EffectivePermit = ProcessAndSafetyPermit combine au couplage synchro (anti-télescopage)
// ET gaté par NOT SafeStop (défauts thermique/phase/codeur/méca) : le permit reflète « prêt à
// fonctionner », aligné sur M3 (PRG_05 §1ter). SafeStopM1/M2_Active agrège déjà le couplage
// synchro (SafeStop de l'autre treuil pendant SyncActive) — cohérent avec l'anti-télescopage.
EffectivePermitM1_Descend := ProcessAndSafetyPermitM1_Descend AND NOT SafeStopM1_Active AND (NOT CoupledBoth OR ProcessAndSafetyPermitM2_Descend);
EffectivePermitM2_Descend := ProcessAndSafetyPermitM2_Descend AND NOT SafeStopM2_Active AND (NOT CoupledBoth OR ProcessAndSafetyPermitM1_Descend);
EffectivePermitM1_Ascent  := ProcessAndSafetyPermitM1_Ascent  AND NOT SafeStopM1_Active AND (NOT CoupledBoth OR ProcessAndSafetyPermitM2_Ascent);
EffectivePermitM2_Ascent  := ProcessAndSafetyPermitM2_Ascent  AND NOT SafeStopM2_Active AND (NOT CoupledBoth OR ProcessAndSafetyPermitM1_Ascent);

// Mode secours MAINT_N2 : pilotage direct inconditionnel des contacteurs M1/M2 (ensemble ou separement)
// sous la seule reserve de la chaine AU physique fermee (PowerContactorEngaged_DI) et du capteur
// mecanique haut (TopPositionFree_DI, sauf bypass explicite).
IF MaintN2 THEN
    SafeStopM1_Active := NOT PRG_02_Acquisition.HwIn.Machine.PowerContactorEngaged_DI;
    SafeStopM2_Active := NOT PRG_02_Acquisition.HwIn.Machine.PowerContactorEngaged_DI;
    EffectivePermitM1_Descend := PRG_02_Acquisition.HwIn.Machine.PowerContactorEngaged_DI;
    EffectivePermitM2_Descend := PRG_02_Acquisition.HwIn.Machine.PowerContactorEngaged_DI;
    EffectivePermitM1_Ascent  := PRG_02_Acquisition.HwIn.Machine.PowerContactorEngaged_DI
                                 AND ((PRG_02_Acquisition.HwIn.Winch.M1M2_TopPositionFree_DI
                                       AND NOT PRG_06_Outputs.Data.TopHardStopLatched)
                                      OR BypassM1TopLimitSwitchEff
                                      OR GVL_IHM.M1TreuilRetenue.Bypass.Global);
    EffectivePermitM2_Ascent  := PRG_02_Acquisition.HwIn.Machine.PowerContactorEngaged_DI
                                 AND ((PRG_02_Acquisition.HwIn.Winch.M1M2_TopPositionFree_DI
                                       AND NOT PRG_06_Outputs.Data.TopHardStopLatched)
                                      OR BypassM2TopLimitSwitchEff
                                      OR GVL_IHM.M2TreuilBenne.Bypass.Global);
END_IF;

// Si un cycle homing machine est actif (en N1 ou N2), appliquer ses permis par etape
IF HomingFreeMoveBlockedN1 THEN
    EffectivePermitM1_Ascent  := FALSE;
    EffectivePermitM1_Descend := FALSE;
    EffectivePermitM2_Ascent  := FALSE;
    EffectivePermitM2_Descend := FALSE;
ELSIF PRG_02_Acquisition.Data.MachineHoming.Active THEN
    IF PRG_02_Acquisition.Data.MachineHoming.CmdWinchSelect = 2 THEN
        EffectivePermitM1_Ascent  := FALSE;
        EffectivePermitM1_Descend := FALSE;
        EffectivePermitM2_Ascent  := EffectivePermitM2_Ascent  AND PRG_02_Acquisition.Data.MachineHoming.AllowAscent;
        EffectivePermitM2_Descend := EffectivePermitM2_Descend AND PRG_02_Acquisition.Data.MachineHoming.AllowDescend;
    ELSIF PRG_02_Acquisition.Data.MachineHoming.CmdWinchSelect = 0 THEN
        EffectivePermitM1_Ascent  := EffectivePermitM1_Ascent  AND PRG_02_Acquisition.Data.MachineHoming.AllowAscent;
        EffectivePermitM1_Descend := EffectivePermitM1_Descend AND PRG_02_Acquisition.Data.MachineHoming.AllowDescend;
        EffectivePermitM2_Ascent  := EffectivePermitM2_Ascent  AND PRG_02_Acquisition.Data.MachineHoming.AllowAscent;
        EffectivePermitM2_Descend := EffectivePermitM2_Descend AND PRG_02_Acquisition.Data.MachineHoming.AllowDescend;
    ELSE
        EffectivePermitM1_Ascent  := FALSE;
        EffectivePermitM1_Descend := FALSE;
        EffectivePermitM2_Ascent  := FALSE;
        EffectivePermitM2_Descend := FALSE;
    END_IF;
END_IF;

// Permis canoniques benne : ouverture = M2 vers le bas, fermeture = M2 vers le haut.
// Les fins de course benne restent des faits fonctionnels distincts des limites treuil.
EffectivePermitBucket_Open := EffectivePermitM2_Descend
    AND PRG_02_Acquisition.Data.EncoderM1.Homed
    AND PRG_02_Acquisition.Data.EncoderM2.Homed
    AND (instBucket.Lifecycle.Busy OR NOT _BucketState.IsOpen)
    AND NOT instBucket.Fault.Error;
EffectivePermitBucket_Close := EffectivePermitM2_Ascent
    AND PRG_02_Acquisition.Data.EncoderM1.Homed
    AND PRG_02_Acquisition.Data.EncoderM2.Homed
    AND (instBucket.Lifecycle.Busy OR NOT _BucketState.IsClosed)
    AND NOT instBucket.Fault.Error;

// Défense en profondeur benne : le permis directionnel benne est appliqué au
// même scan aux deux niveaux M2, uniquement lorsque FB_Bucket est producteur.
M2AscentPermitApplied := EffectivePermitM2_Ascent
    AND (NOT instBucket.M2_RunRequest OR EffectivePermitBucket_Close);
M2DescendPermitApplied := EffectivePermitM2_Descend
    AND (NOT instBucket.M2_RunRequest OR EffectivePermitBucket_Open);

// 🔗 Agrégats Both : permis communs consommés par la commande both.
// = AND des 4 permits effectifs. Chaque axe garde sa vérité propre
// (EffectivePermitM*_*) ; en commande both, seul l'agrégat est consommé (§6),
// garantissant "les 2 treuils partent ensemble, ou aucun".

// 📉 Diagnostic IHM — cause priorisée du blocage Both (lecture seule, NC-100).
// N'a AUCUN effet de conduite : l'arrêt est porté par Both*Permit (§6, consommé par les
// 2 FB_Winch) et la défense en profondeur par la barrière finale (FB_WinchOutputInterlock,
// coupe par PermitFinalBlocked). Ordre : cause la plus grave gagne.
IF NOT WinchBothMotionActive THEN
    BothBlocked             := FALSE;
    BothBlockReason         := E_WinchTraceBlockReason.NONE;
ELSIF NOT ((WinchBothReqAscent AND EffectivePermitM1_Ascent AND EffectivePermitM2_Ascent)
        OR (WinchBothReqDescend AND EffectivePermitM1_Descend AND EffectivePermitM2_Descend)) THEN
    BothBlocked             := TRUE;
    BothBlockReason         := E_WinchTraceBlockReason.COUPLING_BLOCKED;
ELSE
    BothBlocked             := FALSE;
    BothBlockReason         := E_WinchTraceBlockReason.NONE;
END_IF;

// 🛡️ ArmingPermit : armer HONNETEMENT, seulement si au moins une action
// selectionnee peut REELLEMENT partir. Disponibilite par axe x sens + motif de
// blocage decode pour l'IHM / troubleshooting. Reprise apres perte = nouveau front
// homme-mort global (FB_Joystick : IF NOT ArmingPermit -> desarme le geste entier).
// EffectivePermitM*_* couvre deja process + safety + NOT SafeStop de cet axe +
// verif couplage ; on ajoute NOT Fault.Latched (faute finale) et, pour M3, le
// permis effectif directionnel + SafeStop/PowerCutOff M3 (bus PRG_05, lag 1 scan).
ArmM1AscentAvail  := EffectivePermitM1_Ascent  AND (MaintN2 OR NOT instSafetyWinchM1.Fault.Latched);
ArmM1DescendAvail := EffectivePermitM1_Descend AND (MaintN2 OR NOT instSafetyWinchM1.Fault.Latched);
ArmM2AscentAvail  := EffectivePermitM2_Ascent  AND (MaintN2 OR NOT instSafetyWinchM2.Fault.Latched);
ArmM2DescendAvail := EffectivePermitM2_Descend AND (MaintN2 OR NOT instSafetyWinchM2.Fault.Latched);
ArmM3TremieAvail  := PRG_05_Translation.Data.TranslationFinalInterlockRequest.EffectivePermitM3_Tremie
                     AND NOT PRG_05_Translation.Data.TranslationSafety.SafeStop
                     AND NOT PRG_05_Translation.Data.TranslationSafety.PowerCutOff;
ArmM3MaintenanceAvail := PRG_05_Translation.Data.TranslationFinalInterlockRequest.EffectivePermitM3_Maintenance
                     AND NOT PRG_05_Translation.Data.TranslationSafety.SafeStop
                     AND NOT PRG_05_Translation.Data.TranslationSafety.PowerCutOff;

ArmAnyAxisAvail := ArmM1AscentAvail OR ArmM1DescendAvail
               OR ArmM2AscentAvail OR ArmM2DescendAvail
               OR ArmM3TremieAvail OR ArmM3MaintenanceAvail;

// Conditions de base (AC1) — priorite decroissante pour le motif.
// En SEMI_AUTO ou lors d'une commande benne programme (AX3_OPEN_BUCKET / vidage), l'operateur
// doit pouvoir armer l'homme-mort (DeadmanArmed) pour autoriser le mouvement benne !
ArmBucketBusy := (instBucket.Lifecycle.Busy OR BenneBusyFallEdge.Q)
                 AND NOT MaintN2
                 AND NOT PRG_02_Acquisition.Data.MachineHoming.Active
                 AND (PRG_03_Modes_Cycle.Data.Auth.Mode <> E_Mode.SEMI_AUTO)
                 AND NOT PRG_03_Modes_Cycle.Data.ReqProgram.ReqBucket.ReqOpen
                 AND NOT PRG_03_Modes_Cycle.Data.ReqProgram.ReqBucket.ReqClose;
ArmModeDisabled := (PRG_03_Modes_Cycle.Data.Auth.Mode = E_Mode.DISABLE);
ArmContactorOff := NOT PRG_02_Acquisition.HwIn.Machine.PowerContactorEngaged_DI;
ArmPowerCutOff := NOT MaintN2
               AND (instSafetyWinchM1.PowerCutOff OR instSafetyWinchM2.PowerCutOff
                    OR PRG_05_Translation.Data.TranslationSafety.PowerCutOff);

IF ArmModeDisabled THEN
    Data.ArmingAvailability.BlockedReason := E_ArmingBlockReason.MODE_DISABLE;
ELSIF ArmContactorOff THEN
    Data.ArmingAvailability.BlockedReason := E_ArmingBlockReason.CONTACTOR_OFF;
ELSIF ArmPowerCutOff THEN
    Data.ArmingAvailability.BlockedReason := E_ArmingBlockReason.POWER_CUTOFF;
ELSIF ArmBucketBusy THEN
    Data.ArmingAvailability.BlockedReason := E_ArmingBlockReason.BUCKET_BUSY;
ELSIF NOT ArmAnyAxisAvail THEN
    Data.ArmingAvailability.BlockedReason := E_ArmingBlockReason.ALL_AXES_BLOCKED;
ELSE
    Data.ArmingAvailability.BlockedReason := E_ArmingBlockReason.NONE;
END_IF;

ArmingPermit := NOT ArmModeDisabled AND NOT ArmContactorOff AND NOT ArmPowerCutOff
             AND NOT ArmBucketBusy AND ArmAnyAxisAvail;

Data.ArmingAvailability.M1AscentAvail      := ArmM1AscentAvail;
Data.ArmingAvailability.M1DescendAvail     := ArmM1DescendAvail;
Data.ArmingAvailability.M2AscentAvail      := ArmM2AscentAvail;
Data.ArmingAvailability.M2DescendAvail     := ArmM2DescendAvail;
Data.ArmingAvailability.M3TremieAvail      := ArmM3TremieAvail;
Data.ArmingAvailability.M3MaintenanceAvail := ArmM3MaintenanceAvail;
Data.ArmingAvailability.AnyAxisAvail       := ArmAnyAxisAvail;

{endregion}

{region "📐 §5ter Clamp palier"}
// === 🧮 §5ter AGRÉGATEUR DE CLAMP DE PALIER ===
// Bornes communes identiques M1=M2, puis M2 applique ses limites benne propres.
// Plafond = MIN des sources plafond ; plancher = MAX des sources plancher ; plafond gagne.
// Synchro (instWinchSync) calculée en §4, en amont : SyncDeviationWarn réduit les DEUX treuils.

// --- Sources communes (M1 = M2) ---
CommonMaxStepAscent   := EffectiveMaxStepAscent;
CommonMaxStepDescent := EffectiveMaxStepDescent;

// Plafond fixe demandé : en position Maintenance validée par front, les deux
// treuils restent limités au palier 1 dans les deux sens. Ces valeurs ne sont
// volontairement pas exposées comme consignes IHM : une IHM ne doit pas pouvoir
// relever un garde-fou de vitesse.
MaintenanceMaxStepAscent  := 1;
MaintenanceMaxStepDescent := 1;

// SECURITE ISO 13849 - posture fail-safe : bridage vitesse hors homing.
// Codeurs non references => position non fiable => plafond palier 1 sur M1 ET M2,
// montee ET descente. Symetrique (aucun vecteur contacteur M1<>M2). Sans ce garde-fou,
// palier 5 accessible non reference : les caps de position (SlowdownMaxStep,
// SyncDeviationWarn) sont eux-memes inactifs sans reference fiable. Debridage assume
// plus tard sur capteur haut actif (position redevenue connue).
IF PRG_02_Acquisition.Data.MachineHoming.Active
   OR NOT (PRG_02_Acquisition.Data.EncoderM1.HomedAndReliable
           AND PRG_02_Acquisition.Data.EncoderM2.HomedAndReliable) THEN
    CommonMaxStepAscent  := 1;
    CommonMaxStepDescent := 1;
END_IF;

IF instWinchSync.SyncDeviationWarn THEN
    CommonMaxStepAscent   := 1;
    CommonMaxStepDescent := 1;
END_IF;
IF PRG_03_Modes_Cycle.Data.ReqProgram.ReqBucket.ExtractionControlActive OR ExtractionControlActive THEN
    CommonMaxStepAscent := 1;
END_IF;
// Benne non fermee (ou mou de cable) EN PILOTAGE COUPLE : les DEUX treuils a palier 1.
// Brider M2 seul (bloc M2-propre ci-dessous) laisserait M1 monter plus vite -> vecteurs
// contacteurs M1<>M2 -> FB_SyncContactor (PRG_06) -> ContactorMismatch -> SafeStop.
// En couple les 2 treuils sont lies : la limite benne s'applique aux 2.
IF CoupledBoth AND (BucketNotClosedAscentCapStep1 OR SlackCableAscentCapStep1) THEN
    CommonMaxStepAscent := 1;
END_IF;

// En pilotage Both (WinchBothMotionActive), M1 est l'unique autorité nominale
// de vitesse en approche haute. Dès que M1 entre dans sa zone de ralentissement haut,
// CommonMaxStepAscent est bridé à WinchSlowdownMaxStep (palier 1). Cela garantit que M1 et M2
// décélèrent de façon synchrone et atomique au palier 1, éliminant la divergence de paliers
// P1/P5 qui causait une neutralisation brutale sous WinchBothFinalRequestsCoherent.
IF WinchBothMotionActive
   AND PRG_02_Acquisition.Data.EncoderM1.Homed
   AND NOT PRG_02_Acquisition.Data.EncoderM1.HomingSuspect
   AND (PRG_02_Acquisition.Data.EncoderM1.Measurement.CablePosM >= (TopLimitM1_M - _CommunCfgPersist.WinchSlowdownDistanceTop_M)) THEN
    CommonMaxStepAscent := MIN(CommonMaxStepAscent, _CommunCfgPersist.WinchSlowdownMaxStep);
END_IF;

// Position Maintenance atteinte : bridage commun M1/M2, montée et descente.
// Ne pas utiliser SensorsWord ici : il décrit une zone, pas une position validée.
IF PRG_05_Translation.Data.M3_AtMaintenanceStable THEN
    CommonMaxStepAscent  := MIN(CommonMaxStepAscent, MaintenanceMaxStepAscent);
    CommonMaxStepDescent := MIN(CommonMaxStepDescent, MaintenanceMaxStepDescent);
END_IF;

// Planchers communs : 1 (neutre) en montée ; en descente, 0 hors plongée.
// MinStepDown=0 signifie explicitement « aucun plancher » : seul FB_DiveSearch
// peut imposer un palier de plongée. Ne jamais réintroduire un minimum à 1 ici,
// sinon une inversion de sens ne peut plus atteindre StepNumber=0.
// Règle de l'agrégateur : plancher = MAX des sources plancher ; si plancher > plafond,
// LE PLAFOND GAGNE — le clamp final (consommation FB_Winch, lot aval) borne au plafond,
// on ne force donc jamais ici un palier au-delà de CommonMaxStepDescent.
CommonMinStepUp   := 1;
CommonMinStepDown := MAX(0, PRG_03_Modes_Cycle.Data.ReqProgram.ReqBucket.MinStepDown);

// --- M2-propre (jamais vu par M1) ---
M2MaxStepUp   := CommonMaxStepAscent;
M2MaxStepDown := CommonMaxStepDescent;
// T291-A : le plafond nominal commun reste configure a 4 afin que M1 et tous
// les autres modes restent inchanges. Pendant la seule plongee auto AX4..AX7,
// M2 peut atteindre P5. Ne jamais relever ici un plafond deja reduit par une
// protection amont (codeurs non fiables, ecart synchro, position maintenance).
IF PRG_03_Modes_Cycle.Data.AutoDiveM1Step4M2Step5Active
   AND (EffectiveMaxStepDescent = 4)
   AND (CommonMaxStepDescent = EffectiveMaxStepDescent) THEN
    M2MaxStepDown := 5;
END_IF;
// Auto-séquencement benne : AX10 SEMI_AUTO garde le plafond AX11 P1..P2 ; les
// autres manoeuvres benne conservent leur plafond dédié.
IF instBucket.M2_BucketJogLimit THEN
    IF ArbContext.BucketHandoffP1Active THEN
        M2MaxStepUp := 1;
    ELSIF ArbContext.BucketAutoCloseActive THEN
        M2MaxStepUp := MIN(M2MaxStepUp, LIMIT(1, GVL_IHM.CycleSemiAuto.Cfg.CtrlAscentMaxStep, 2));
    ELSE
        M2MaxStepUp := LIMIT(1, _BucketCfgPersist.Config.MaxStepUp, 5);
    END_IF;
    M2MaxStepDown := LIMIT(1, _BucketCfgPersist.Config.MaxStepDown, 5);
END_IF;
// Jog unitaire M2 : palier libre en course, palier 1 uniquement dans la zone de
// ralentissement (JogSlowdownZoneM avant le point d'arrêt anticipé — cf. §5). Montée M2
// = fermeture, descente M2 = ouverture. Les zones sont calculées sur la position :
// si M1/M2 ne sont pas référencés, la position n'a pas de sens → repli palier 1 partout.
IF ManualBucketJogActive THEN
    IF PRG_02_Acquisition.Data.MachineHoming.Active
       OR NOT (PRG_02_Acquisition.Data.EncoderM1.Homed AND PRG_02_Acquisition.Data.EncoderM2.Homed) THEN
        M2MaxStepUp   := 1;
        M2MaxStepDown := 1;
    ELSE
        M2MaxStepUp   := MIN(M2MaxStepUp, LIMIT(1, _BucketCfgPersist.Config.MaxStepUp, 5));
        M2MaxStepDown := MIN(M2MaxStepDown, LIMIT(1, _BucketCfgPersist.Config.MaxStepDown, 5));
        IF M2JogApproachClose THEN
            M2MaxStepUp := 1;
        END_IF;
        IF M2JogApproachOpen THEN
            M2MaxStepDown := 1;
        END_IF;
    END_IF;
END_IF;
IF SlackCableAscentCapStep1
   OR (BucketNotClosedAscentCapStep1 AND NOT ArbContext.BucketAutoCloseActive) THEN
    M2MaxStepUp := 1;
END_IF;

// Protection finale M2 : les limites spécifiques benne ne peuvent pas remonter
// le plafond fixe de sécurité appliqué en position Maintenance.
IF PRG_05_Translation.Data.M3_AtMaintenanceStable THEN
    M2MaxStepUp   := MIN(M2MaxStepUp, MaintenanceMaxStepAscent);
    M2MaxStepDown := MIN(M2MaxStepDown, MaintenanceMaxStepDescent);
END_IF;
M2MinStepUp   := CommonMinStepUp;
M2MinStepDown := CommonMinStepDown;
{endregion}

{region "⚙️ §6 Exécution M1/M2"}
// === ⚙️ §6 EXÉCUTION FB_Winch (M1 & M2) ===

// Estimateurs de bande vitesse réelle appelés AVANT instWinchM1/M2 : leur sortie
// SpeedBand alimente MeasuredSpeedBand (2e étage du garde-fou FB_Winch) sur le même
// scan. Sources vitesse identiques à FB_Safety_Winch (§5bis).
instWinchLoadEstimatorM1(
    Enable                  := (PRG_03_Modes_Cycle.Data.Auth.Mode <> E_Mode.DISABLE) AND NOT PRG_03_Modes_Cycle.Data.Auth.InhibitM1,
    Reset                   := PRG_07_Supervision.FaultMachineReset_IHM,
    Mode                    := PRG_03_Modes_Cycle.Data.Auth.Mode,
    ActiveSpeedStep         := instWinchM1.StepNumber,
    PowerContactorEngaged   := PRG_02_Acquisition.HwIn.Machine.PowerContactorEngaged_DI,
    MeasuredSpeedMps        := PRG_02_Acquisition.Data.EncoderM1.Measurement.Speed_Mps,
    MeasuredSpeedSignedMps  := PRG_02_Acquisition.Data.EncoderM1.Measurement.SignedSpeed_Mps,
    SpeedConfig             := _WinchSpeedConfig,
    LoadTable               := _WinchLoadEstimateTable
);

instWinchLoadEstimatorM2(
    Enable                  := (PRG_03_Modes_Cycle.Data.Auth.Mode <> E_Mode.DISABLE) AND NOT PRG_03_Modes_Cycle.Data.Auth.InhibitM2,
    Reset                   := PRG_07_Supervision.FaultMachineReset_IHM,
    Mode                    := PRG_03_Modes_Cycle.Data.Auth.Mode,
    ActiveSpeedStep         := instWinchM2.StepNumber,
    PowerContactorEngaged   := PRG_02_Acquisition.HwIn.Machine.PowerContactorEngaged_DI,
    MeasuredSpeedMps        := PRG_02_Acquisition.Data.EncoderM2.Measurement.Speed_Mps,
    MeasuredSpeedSignedMps  := PRG_02_Acquisition.Data.EncoderM2.Measurement.SignedSpeed_Mps,
    SpeedConfig             := _WinchSpeedConfig,
    LoadTable               := _WinchLoadEstimateTable
);

// --- M1 : assemblage des structs (CODESYS refuse l'initialiseur inline en appel) ---
// 🔗 Routage permit both : en commande both (WinchBothMotionActive=TRUE), les
// Chaque treuil consomme directement son permis directionnel canonique ; Both est
// validé par l'AND des deux axes dans l'arbitrage.
// jamais les permits individuels directement. En unitaire (M1 seul / M2 seul / benne M2),
// chacun consomme son permit effectif propre (comportement inchangé). SEL(a, b, c) := a ? c : b.
ReqM1Winch.RunRequest               := M1LogicRunRequest;
ReqM1Winch.ReqAscent                := M1LogicReqAscent;
ReqM1Winch.ReqDescend               := M1LogicReqDescend;
ReqM1Winch.SpeedStepReq             := M1LogicRequestStepTgt;

// === ATOMICITE DU DEMARRAGE COUPLE (verrou boucle fermee, remplace le timer aveugle) ===
// En intention both (WinchSel=0), TANT QU'un des deux treuils n'est pas pret a bouger
// -- encore dans son dead-time D18 (FB_WinchDirectionInterlock, arme apres un arret, ex.
// fin de jog benne) OU en defaut latche -- on FIGE la commande FINALE des DEUX. Le treuil
// qui vient de s'arreter garde ainsi son delai en cours ; quand il est pret, les deux
// contacteurs s'enclenchent au MEME cycle -> 0 cm de decalage tambours (REX MES 2026-09-04 :
// M1 parti seul 59 cm apres ouverture benne). instWinchM2.* = valeur du scan precedent
// (lag 1 scan assume : la garde tient juste 1 scan de plus, sans risque).
//
// REGLE : on fige UNIQUEMENT le treuil PRET, jamais celui qui purge son dead-time.
// Zeroter la requete d'un treuil efface son propre DeadTimeArmed (NOT RequestActive) ->
// si on figeait les deux, M2 perdrait son delai D18 et la garde s'effondrerait en 1 scan.
// Donc : M1 pret + M2 en dead-time -> on fige M1, on laisse M2 finir son delai ; au scan
// ou M2 devient pret, les deux demarrent ensemble.
WinchBothMotionReady := NOT (instWinchM1.DirectionChangePending OR instWinchM2.DirectionChangePending)
                        AND NOT instWinchM1.Fault.Latched AND NOT instWinchM2.Fault.Latched;
IF NOT MaintN2 AND WinchBothMotionActive AND (instWinchM2.DirectionChangePending OR instWinchM2.Fault.Latched) THEN
    ReqM1Winch.RunRequest := FALSE; ReqM1Winch.ReqAscent := FALSE; ReqM1Winch.ReqDescend := FALSE; ReqM1Winch.SpeedStepReq := 0;
END_IF;
ReqM1Winch.MaxStepUp                := CommonMaxStepAscent;
ReqM1Winch.MaxStepDown              := CommonMaxStepDescent;
// Plancher palier descente plongée Kobold : plancher plongée agrégé en §5ter, injecté
// sur la cible (jamais sur StepNumber). Aucun effet si StartStop=FALSE.
ReqM1Winch.MinStepDown              := CommonMinStepDown;
ReqM1Winch.HomingApproachActive     := PRG_03_Modes_Cycle.Data.Auth.HomingApproachEnable;
// Même limite haute active que FB_Safety_Winch (7,5 m / 8,5 m sous override).
ReqM1Winch.TopLimitM                := TopLimitM1_M;
ReqM1Winch.BottomLimitM             := BottomLimitM1_Active;
ReqM1Winch.SyncCoupled              := instWinchSync.SyncActive;
